               IF #Kamera.text_etiketa = '' THEN
                   #Kamera.text_etiketa := 'NECTENO';   // prazdny text = prazdna pozice!
               END_IF;

               // zapis ZA posledni obsazenou pozici
               #Kamera.idx := 0;
               FOR #i := 5 TO 1 BY -1 DO
                   IF "DB_HMI_recype".fronta[#i].prenaseny_text <> '' THEN
                       #Kamera.idx := #i;
                       EXIT;
                   END_IF;
               END_FOR;

               IF #Kamera.idx < 5 THEN
                   "DB_HMI_recype".fronta[#Kamera.idx + 1].prenaseny_text := #Kamera.text_etiketa;
                   "DB_HMI_recype".fronta[#Kamera.idx + 1].balik_den := #Kamera.balik_den;
                   "DB_HMI_recype".fronta[#Kamera.idx + 1].vyrazeni := #Kamera.vyradit;
               ELSE
                   #Kamera.fronta_plna := TRUE;
               END_IF;
               #Kamera.sber_aktivni := FALSE;
           END_IF;
       END_REGION

       REGION Novy balik pod kamerou - start sberu (az PO zapisu predchoziho)
           IF #Kamera.s2_nabeh THEN
               // citac plat (presunuto ze site 20)
               #zpracovani_dat[1].balik_den := #zpracovani_dat[1].balik_den + 1;
               IF #zpracovani_dat[1].balik_den >= 32000 THEN
                   #zpracovani_dat[1].balik_den := 1;
               END_IF;
               #Kamera.balik_den := #zpracovani_dat[1].balik_den;   // az PO pricteni

               #Kamera.sber_aktivni := TRUE;
               #Kamera.prijato_etiketa := FALSE;
               #Kamera.prijato_folie_l := FALSE;
               #Kamera.prijato_folie_p := FALSE;
               #Kamera.ok_etiketa := FALSE;
               #Kamera.ok_folie_l := FALSE;
               #Kamera.ok_folie_p := FALSE;
               #Kamera.text_etiketa := '';
           END_IF;
       END_REGION
   END_IF;

   REGION Obsazenost fronty pro HMI (pocita se kazdy scan)
       #Kamera.pocet := 0;
       FOR #i := 1 TO 5 DO
           IF "DB_HMI_recype".fronta[#i].prenaseny_text <> '' THEN
               #Kamera.pocet := #Kamera.pocet + 1;
           END_IF;
       END_FOR;
       "DB_HMI_recype".obsazenost_fronty := #Kamera.pocet;
       IF #Kamera.pocet = 0 THEN
           #Kamera.fronta_plna := FALSE;
       END_IF;
   END_REGION
END_REGION

REGION Network 22 (SCL): PŘEPNUTÍ JOBU HORNÍ KAMERY
   // Prepnuti jobu horni kamery podle receptury.
   // Spousti se nabeznou hranou "DB_HMI_recype".ODESLI_dATA (tlacitko Odeslani dat do tiskarny)
   // - soubezne s odeslanim zpravy do tiskarny (OP2).
   // Job 0 v recepture = job neprepinat.

   #Kam_Etiketa_Job.pozadovany := "DB_HMI_recype".recipe.PRG_CAM_etiketa;

   IF "CONTROL_LINE_DB".trig.reset_error_all THEN
       #Kam_Etiketa_Job.chyba := FALSE;
   END_IF;

   CASE #Kam_Etiketa_Job.krok OF
       0:  // ---- klid: cekam na pozadavek ----
           #Kam_Etiketa_Job.aktivni := FALSE;
           "COG_ETIKETA_is3800-ExecuteCommand/JobLoad" := FALSE;
           IF "DB_HMI_recype".ODESLI_dATA AND NOT #Kam_Etiketa_Job.odesli_pamet
               AND #Kam_Etiketa_Job.pozadovany > 0
               AND "COG_ETIKETA_is3800-Online" THEN
               "COG_ETIKETA_is3800-CommandID" := INT_TO_WORD(#Kam_Etiketa_Job.pozadovany);
               #Kam_Etiketa_Job.aktivni := TRUE;
               #Kam_Etiketa_Job.chyba := FALSE;
               #Kam_Etiketa_Job.krok := 10;
           END_IF;

       10: // ---- CommandID uz je venku (predchozi cyklus) -> spustit prikaz ----
           "COG_ETIKETA_is3800-ExecuteCommand/JobLoad" := TRUE;
           #Kam_Etiketa_Job.krok := 20;

       20: // ---- cekam na vysledek ----
           IF "COG_ETIKETA_is3800-CommandCompleted" THEN
               #Kam_Etiketa_Job.krok := 30;
           ELSIF "COG_ETIKETA_is3800-CommandFailed" THEN
               #Kam_Etiketa_Job.chyba := TRUE;
               #Kam_Etiketa_Job.chyba_kod := "COG_ETIKETA_is3800-CommandResultCode";
               #Kam_Etiketa_Job.krok := 30;
           ELSIF #TIMER.TIMER_3.Q THEN
               #Kam_Etiketa_Job.chyba := TRUE;            // kamera neodpovedela
               #Kam_Etiketa_Job.chyba_kod := 16#FFFF;
               #Kam_Etiketa_Job.krok := 30;
           END_IF;

       30: // ---- ukonceni handshake: shodit Execute, pockat az kamera shodi stav ----
           "COG_ETIKETA_is3800-ExecuteCommand/JobLoad" := FALSE;
           IF NOT "COG_ETIKETA_is3800-CommandCompleted"
               AND NOT "COG_ETIKETA_is3800-CommandFailed" THEN
               #Kam_Etiketa_Job.krok := 0;
           END_IF;

       ELSE
           #Kam_Etiketa_Job.krok := 0;
   END_CASE;

   // casovac timeoutu bezi v krocich 10..30
   #TIMER.TIMER_3.TON(IN := #Kam_Etiketa_Job.krok >= 10,
                      PT := #Kam_Etiketa_Job.timeout);
   IF #TIMER.TIMER_3.Q AND #Kam_Etiketa_Job.krok = 30 THEN
       #Kam_Etiketa_Job.krok := 0;                         // pojistka, kdyby kamera stav neshodila
   END_IF;

   #Kam_Etiketa_Job.odesli_pamet := "DB_HMI_recype".ODESLI_dATA;

   // kontrola: v klidu musi job v kamere odpovidat recepture
   #Kam_Etiketa_Job.nesouhlasi := #Kam_Etiketa_Job.krok = 0
   AND #Kam_Etiketa_Job.pozadovany > 0
   AND "COG_ETIKETA_is3800-Online"
   AND WORD_TO_INT("COG_ETIKETA_is3800-Current Job ID") <> #Kam_Etiketa_Job.pozadovany;
END_REGION

REGION Network 23: EXTERNAL_TRIGER
   RUNG wire#powerrail
      { S7_Templates := "SrcType := Int" } EQ_Contact(in1 := #SQCR, in2 := #STEP_5_HOME)
      Contact( "INICIALIZACE_RUN" )
      I_Contact( #TRIG.inicial_ok_op )
      Contact( "AUTOMAT" )
      S_Coil( #HMI.reset_fronty )
      S_Coil( #TRIG.inicial_ok_op )
   END_RUNG
   RUNG wire#powerrail
      Contact( "FirstScan" )
      S_Coil( #HMI.reset_fronty )
      Move(in := 0, out1 => "DB_HMI_recype".obsazenost_fronty, out2 => #zpracovani_dat[1].balik_den)
   END_RUNG
   // the same network as SCL:
   IF (#SQCR = #STEP_5_HOME) AND "INICIALIZACE_RUN" AND NOT #TRIG.inicial_ok_op AND "AUTOMAT" THEN
       #HMI.reset_fronty := TRUE;
       #TRIG.inicial_ok_op := TRUE;
   END_IF;
   IF "FirstScan" THEN
       #HMI.reset_fronty := TRUE;
       "DB_HMI_recype".obsazenost_fronty := 0;
       #zpracovani_dat[1].balik_den := 0;
   END_IF;
END_REGION

REGION Network 24: ETERNAL_TRIGR_INICIAL
   RUNG wire#powerrail
      Contact( "AUTOMAT" )
      { S7_Templates := "SrcType := Int" } GT_Contact(in1 := #SQCR, in2 := #STEP_0)
      { S7_Templates := "SrcType := Int" } LT_Contact(in1 := #SQCR, in2 := #STEP_1000)
      I_Contact( #Kam_Etiketa_Job.aktivni )
      Coil( "COG_ETIKETA_COG_ETIKETA_is3800-TriggerEnable" )
   END_RUNG
   RUNG wire#powerrail
      Contact( "AUTOMAT" )
      { S7_Templates := "SrcType := Int" } GT_Contact(in1 := #SQCR, in2 := #STEP_0)
      { S7_Templates := "SrcType := Int" } LT_Contact(in1 := #SQCR, in2 := #STEP_1000)
      Coil( "COG_FOLIE_L_COG_FOLIE_L_is3800-TriggerEnable" )
   END_RUNG
   RUNG wire#powerrail
      Contact( "AUTOMAT" )
      { S7_Templates := "SrcType := Int" } GT_Contact(in1 := #SQCR, in2 := #STEP_0)
      { S7_Templates := "SrcType := Int" } LT_Contact(in1 := #SQCR, in2 := #STEP_1000)
      Coil( "COG_FOLIE_P_COG_FOLIE_P_is3800-TriggerEnable" )
   END_RUNG
   // the same network as SCL:
   "COG_ETIKETA_COG_ETIKETA_is3800-TriggerEnable" := "AUTOMAT" AND (#SQCR > #STEP_0) AND (#SQCR < #STEP_1000) AND NOT #Kam_Etiketa_Job.aktivni;
   "COG_FOLIE_L_COG_FOLIE_L_is3800-TriggerEnable" := "AUTOMAT" AND (#SQCR > #STEP_0) AND (#SQCR < #STEP_1000);
   "COG_FOLIE_P_COG_FOLIE_P_is3800-TriggerEnable" := "AUTOMAT" AND (#SQCR > #STEP_0) AND (#SQCR < #STEP_1000);
END_REGION

REGION Network 25: hmi
END_REGION

REGION Network 26 (SCL): VYRAZENI MANUAL
   (* #Test_tp_ka12(IN := "DB_Manual".test_vyr,
                 PT := T#500MS);

   "-KA12" := #Test_tp_ka12.Q;

   // testovací bit se sám shodí → každý Modify TRUE = jeden pulz
   IF "DB_Manual".test_vyr THEN
       "DB_Manual".test_vyr := FALSE;
   END_IF; *)
END_REGION
END_FUNCTION_BLOCK

FUNCTION_BLOCK "OP2"   // FB51, LAD
{ S7_Optimized_Access := 'FALSE' }
VERSION : 0.1
   VAR
      CONTROL_MAN : Struct
         B0 : Bool;
         B1 : Bool;
         B2 : Bool;
         B3 : Bool;
         B4 : Bool;
         B5 : Bool;
         B6 : Bool;
         B7 : Bool;
         B8 : Bool;
         B9 : Bool;
         odfuk_1 : Bool;
         odfuk_2 : Bool;
         B12 : Bool;
         B13 : Bool;
         B14 : Bool;
         B15 : Bool;
         B16 : Bool;
         B17 : Bool;
         B18 : Bool;
         B19 : Bool;
         B20 : Bool;
         B21 : Bool;
         B22 : Bool;
         B23 : Bool;
         B24 : Bool;
         B25 : Bool;
         B26 : Bool;
         B27 : Bool;
         B28 : Bool;
         B29 : Bool;
         B30 : Bool;
         B31 : Bool;
      END_STRUCT;
      CONTROL_AUTOMAT : Struct
         connect : Bool;
         send : Bool;
         reciv : Bool;
         trcv : Bool;
         discon : Bool;
         B5 : Bool;
         B6 : Bool;
         B7 : Bool;
         B8 : Bool;
         B9 : Bool;
         B10 : Bool;
         B11 : Bool;
         B12 : Bool;
         B13 : Bool;
         B14 : Bool;
         B15 : Bool;
         B16 : Bool;
         B17 : Bool;
         B18 : Bool;
         B19 : Bool;
         B20 : Bool;
         B21 : Bool;
         B22 : Bool;
         B23 : Bool;
         B24 : Bool;
         B25 : Bool;
         B26 : Bool;
         B27 : Bool;
         B28 : Bool;
         B29 : Bool;
         B30 : Bool;
         B31 : Bool;
      END_STRUCT;
      SENSORS : Struct
         S0 : Bool;
         S1 : Bool;
         S2 : Bool;
         S3 : Bool;
         S4 : Bool;
         S5 : Bool;
         S6 : Bool;
         S7 : Bool;
         S8 : Bool;   // KARUSEL JE NATOČEN PŘÍPRAVKEM A K BRÁNĚ
         S9 : Bool;
         S10 : Bool;
         S11 : Bool;
         S12 : Bool;
         S13 : Bool;
         S14 : Bool;
         S15 : Bool;
         S16 : Bool;
         S17 : Bool;
         S18 : Bool;
         S19 : Bool;
         S20 : Bool;
         S21 : Bool;
         S22 : Bool;
         S23 : Bool;
         S24 : Bool;
         S25 : Bool;
         S26 : Bool;
         S27 : Bool;
         S28 : Bool;
         S29 : Bool;
         S30 : Bool;
         S31 : Bool;
      END_STRUCT;
      SENSORS_1 : Struct
         S0 : Bool;
         S1 : Bool;
         S2 : Bool;
         S3 : Bool;
         S4 : Bool;
         S5 : Bool;
         S6 : Bool;
         S7 : Bool;
         S8 : Bool;
         S9 : Bool;
         S10 : Bool;
         S11 : Bool;
         S12 : Bool;
         S13 : Bool;
         S14 : Bool;
         S15 : Bool;
         S16 : Bool;
         S17 : Bool;
         S18 : Bool;
         S19 : Bool;
         S20 : Bool;
         S21 : Bool;
         S22 : Bool;
         S23 : Bool;
         S24 : Bool;
         S25 : Bool;
         S26 : Bool;
         S27 : Bool;
         S28 : Bool;
         S29 : Bool;
         S30 : Bool;
         S31 : Bool;
      END_STRUCT;
      S_0 : "SENSOR";
      S_1 : "SENSOR";
      S_2 : "SENSOR";
      S_3 : "SENSOR";
      S_4 : "SENSOR";
      S_5 : "SENSOR";
      S_6 : "SENSOR";
      S_7 : "SENSOR";
      S_8 : "SENSOR";
      S_9 : "SENSOR";
      S_10 : "SENSOR";
      S_11 : "SENSOR";
      S_12 : "SENSOR";
      S_13 : "SENSOR";
      S_14 : "SENSOR";
      S_15 : "SENSOR";
      S_16 : "SENSOR";
      M_1 : "MOTOR_CONTROL_BLOCK";
      M_2 : "MOTOR_CONTROL_BLOCK";
      M_3 : "MOTOR_CONTROL_BLOCK";
      SQCR : Int;
      hmi_sqcr : Int;
      TRIG : Struct
         inicial_ok_op : Bool;
         T2 : Bool;
         T3 : Bool;
         T4 : Bool;
         T5 : Bool;
         T6 : Bool;
         T7 : Bool;
         T8 : Bool;
         T9 : Bool;
         T10 : Bool;
         T11 : Bool;
         T12 : Bool;
         T13 : Bool;
         T14 : Bool;
         T15 : Bool;
         T16 : Bool;
         op_1_ready : Bool;
      END_STRUCT;
      MEMOR : Struct
         n_trig_vypnuti : Bool;
         M1 : Bool;
         M2 : Bool;
         M3 : Bool;
         M4 : Bool;
         p_trig_odavacka : Bool;
         M6 : Bool;
         M7 : Bool;
         M8 : Bool;
         M9 : Bool;
         M10 : Bool;
         M11 : Bool;
         RESET_ERROR : Bool;
         M13 : Bool;
         M14 : Bool;
         M15 : Bool;
         SETOVANI_START : Bool;
         M17 : Bool;
         M18 : Bool;
         M19 : Bool;
         M20 : Bool;
         M21 : Bool;
         M22 : Bool;
         M23 : Bool;
         M24 : Bool;
         M25 : Bool;
         M26 : Bool;
         M27 : Bool;
         M28 : Bool;
         M29 : Bool;
         M30 : Bool;
         N_TRIG_SAFETY : Bool;
         M32 : Bool;
         M33 : Bool;
         start_caklu : Bool;
         M35 : Bool;
         M36 : Bool;
         M37 : Bool;
         M38 : Bool;
         M39 : Bool;
         ALARM_GLOBAL : Bool;
         M41 : Bool;
         M42 : Bool;
         M43 : Bool;
         M44 : Bool;
         M45 : Bool;
         M46 : Bool;
         M47 : Bool;
         M48 : Bool;
         M49 : Bool;
         wrong_p_trig : Bool;
         alarm_p_trig : Bool;
         M52 : Bool;
         M53 : Bool;
         M54 : Bool;
         M55 : Bool;
         M56 : Bool;
         M57 : Bool;
         M58 : Bool;
         M59 : Bool;
         M60 : Bool;
         M61 : Bool;
         M62 : Bool;
         M63 : Bool;
      END_STRUCT;
      "TIMER" : Struct
         TIMER_0 : IEC_TIMER;
         TIMER_1 : IEC_TIMER;
         TIMER_2 : IEC_TIMER;
         TIMER_3 : IEC_TIMER;
         TIMER_4 : IEC_TIMER;
         air : IEC_TIMER;
         TIMER_6 : IEC_TIMER;
         TIMER_7 : IEC_TIMER;
      END_STRUCT;
      HMI : Struct
         povoleni_volby_receptu : Bool;
         "svetlo_on/off" : Bool;
         ALARM_VIDITELNOST : Bool;
         hmi_3 : Bool;
         hmi_4 : Bool;
         hmi_5 : Bool;
         hmi_6 : Bool;
         hmi_7 : Bool;
         hmi_8 : Bool;
         hmi_9 : Bool;
         hmi_10 : Bool;
         hmi_11 : Bool;
         hmi_12 : Bool;
         hmi_13 : Bool;
         hmi_14 : Bool;
         hmi_15 : Bool;
      END_STRUCT;
      int_hodnota_zpravy : Word;
      array_do_db AT int_hodnota_zpravy : Array[1..2] of Byte;
      CTRV_LEN : UDInt;
      TCON_Instance : TCON;
      TSEND_Instance : TSEND;
      TRCV_Instance : TRCV;
      TDISCON_Instance : TDISCON;
      Tisk : Struct
         pole2_index_bajt : Int := 14;   // bajt rámce s číslem proměnné
         pole2_index_hodnota : Byte := 16#1;   // číslo proměnné pole 2 (pole 1 = 0)
         datum_chyba : Bool;   // datum přepsáno na XX.XX.XXXX
         pole2_kratky : Bool := true;
         jeden_ramec : Bool;
      END_STRUCT;
   END_VAR
   VAR_TEMP
      DATA : Array[0..255] of Char;
      ARRAY_NULL : Array[1..8] of Bool;
      ARRAY_PRAZDNE : Array[0..255] of Byte;
      j : Int;
      L1 : Int;
      p : Int;
   END_VAR
   VAR CONSTANT
      STEP_0 : Int := 0;
      step_2 : Int := 2;
      STEP_4 : Int := 4;
      STEP_5_HOME : Int := 5;
      STEP_7 : Int := 7;
      STEP_10 : Int := 10;
      STEP_15 : Int := 15;
      STEP_20 : Int := 20;
      STEP_23 : Int := 23;
      STEP_25 : Int := 25;
      STEP_27 : Int := 27;
      STEP_30 : Int := 30;
      STEP_35 : Int := 35;
      STEP_37 : Int := 37;
      STEP_40 : Int := 40;
      STEP_43 : Int := 43;
      STEP_45 : Int := 45;
      STEP_50 : Int := 50;
      STEP_55 : Int := 55;
      STEP_60 : Int := 60;
      STEP_65 : Int := 65;
      STEP_70 : Int := 70;
      STEP_73 : Int := 73;
      STEP_75 : Int := 75;
      STEP_80 : Int := 80;
      STEP_83 : Int := 83;
      STEP_85 : Int := 85;
      STEP_90 : Int := 90;
      STEP_93 : Int := 93;
      STEP_95 : Int := 95;
      STEP_100 : Int := 100;
      STEP_105 : Int := 105;
      STEP_110 : Int := 110;
      STEP_113 : Int := 113;
      STEP_115 : Int := 115;
      STEP_120 : Int := 120;
      STEP_125 : Int := 125;
      STEP_130 : Int := 130;
      STEP_135 : Int := 135;
      STEP_140 : Int := 140;
      STEP_145 : Int := 145;
      STEP_150 : Int := 150;
      STEP_155 : Int := 155;
      STEP_1000 : Int := 1000;
      STEP_1001 : Int := 1001;
      STEP_1002 : Int := 1002;
      STEP_1003 : Int := 1003;
      STEP_1004 : Int := 1004;
      STEP_1005 : Int := 1005;
      STEP_1010 : Int := 1010;
      STEP_1015 : Int := 1015;
      STEP_1020 : Int := 1020;
      STEP_1025 : Int := 1025;
      STEP_3000 : Int := 3000;
      STEP_3005 : Int := 3005;
      STEP_3010 : Int := 3010;
      STEP_3015 : Int := 3015;
      STEP_3020 : Int := 3020;
      STEP_2000 : Int := 2000;
      string_null : String;
      char_null : Char;
      text_kartacek : String := 'Kartacek';
      string_kar_A : String := 'A';
      string_kar_B : String := 'B';
   END_VAR
   VAR_TEMP   // added for the SCL form of the ladder/FBD networks
      _w1 : Bool;
      _w2 : Bool;
      _w3 : Bool;
   END_VAR
BEGIN

REGION Network 1: manuali ovladani reset
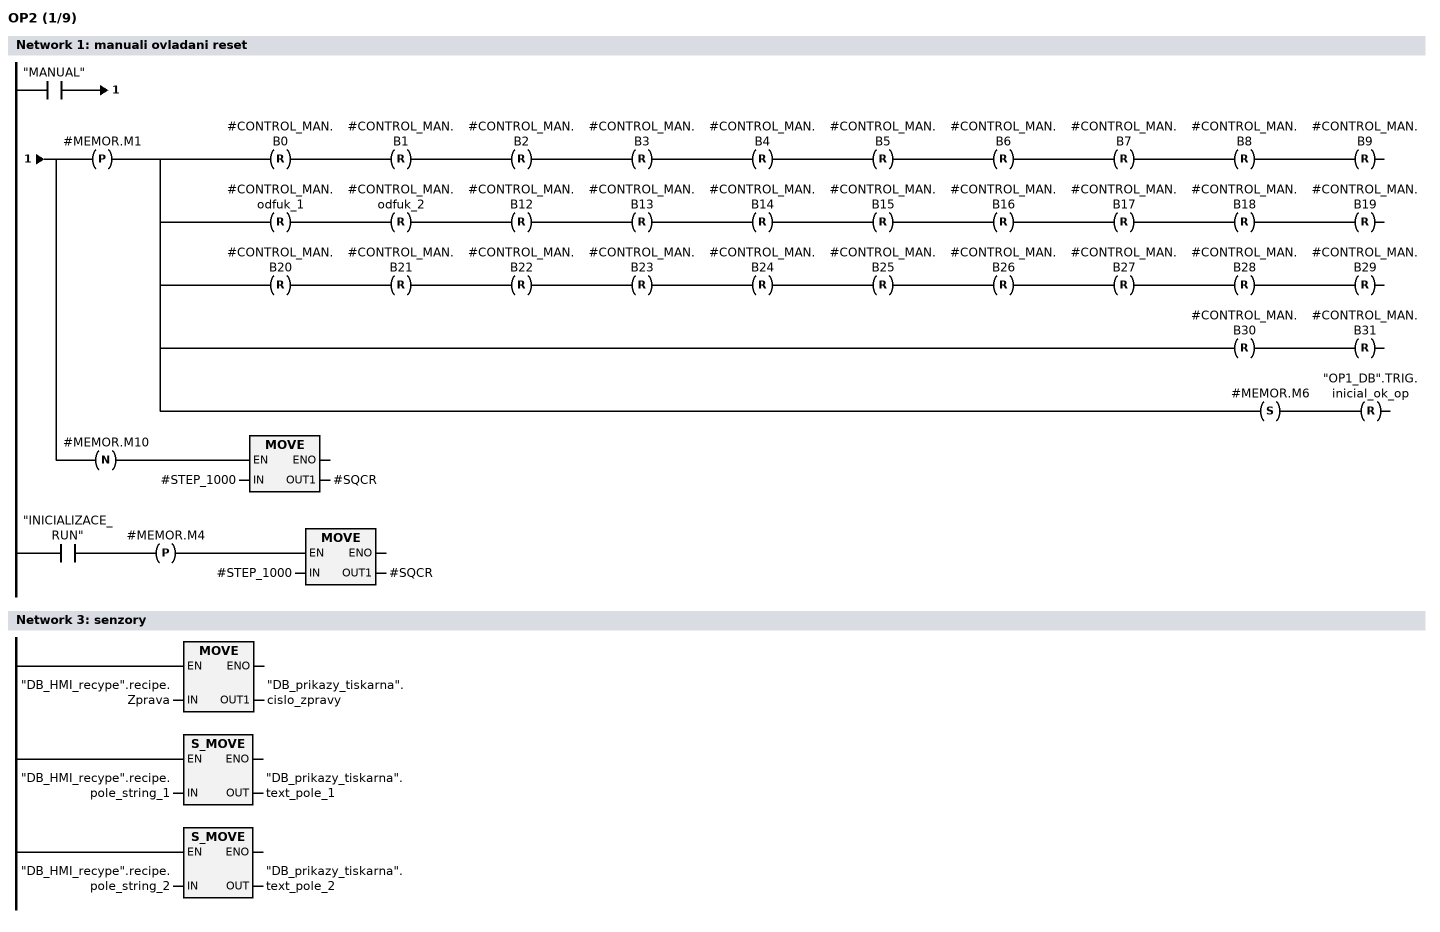
   RUNG wire#powerrail
      Contact( "MANUAL" )
      wire#w1
      P_Trig( #MEMOR.M1 )
      wire#w2
      R_Coil( #CONTROL_MAN.B0 )
      R_Coil( #CONTROL_MAN.B1 )
      R_Coil( #CONTROL_MAN.B2 )
      R_Coil( #CONTROL_MAN.B3 )
      R_Coil( #CONTROL_MAN.B4 )
      R_Coil( #CONTROL_MAN.B5 )
      R_Coil( #CONTROL_MAN.B6 )
      R_Coil( #CONTROL_MAN.B7 )
      R_Coil( #CONTROL_MAN.B8 )
      R_Coil( #CONTROL_MAN.B9 )
   END_RUNG
   RUNG wire#w2
      R_Coil( #CONTROL_MAN.odfuk_1 )
      R_Coil( #CONTROL_MAN.odfuk_2 )
      R_Coil( #CONTROL_MAN.B12 )
      R_Coil( #CONTROL_MAN.B13 )
      R_Coil( #CONTROL_MAN.B14 )
      R_Coil( #CONTROL_MAN.B15 )
      R_Coil( #CONTROL_MAN.B16 )
      R_Coil( #CONTROL_MAN.B17 )
      R_Coil( #CONTROL_MAN.B18 )
      R_Coil( #CONTROL_MAN.B19 )
   END_RUNG
   RUNG wire#w2
      R_Coil( #CONTROL_MAN.B20 )
      R_Coil( #CONTROL_MAN.B21 )
      R_Coil( #CONTROL_MAN.B22 )
      R_Coil( #CONTROL_MAN.B23 )
      R_Coil( #CONTROL_MAN.B24 )
      R_Coil( #CONTROL_MAN.B25 )
      R_Coil( #CONTROL_MAN.B26 )
      R_Coil( #CONTROL_MAN.B27 )
      R_Coil( #CONTROL_MAN.B28 )
      R_Coil( #CONTROL_MAN.B29 )
   END_RUNG
   RUNG wire#w2
      R_Coil( #CONTROL_MAN.B30 )
      R_Coil( #CONTROL_MAN.B31 )
   END_RUNG
   RUNG wire#w2
      S_Coil( #MEMOR.M6 )
      R_Coil( "OP1_DB".TRIG.inicial_ok_op )
   END_RUNG
   RUNG wire#w1
      N_Trig( #MEMOR.M10 )
      Move(in := #STEP_1000, out1 => #SQCR)
   END_RUNG
   RUNG wire#powerrail
      Contact( "INICIALIZACE_RUN" )
      P_Trig( #MEMOR.M4 )
      Move(in := #STEP_1000, out1 => #SQCR)
   END_RUNG
   // the same network as SCL:
   #_w1 := "MANUAL" AND NOT #MEMOR.M1;   // rising edge
   #MEMOR.M1 := "MANUAL";
   IF #_w1 THEN
       #CONTROL_MAN.B0 := FALSE;
       #CONTROL_MAN.B1 := FALSE;
       #CONTROL_MAN.B2 := FALSE;
       #CONTROL_MAN.B3 := FALSE;
       #CONTROL_MAN.B4 := FALSE;
       #CONTROL_MAN.B5 := FALSE;
       #CONTROL_MAN.B6 := FALSE;
       #CONTROL_MAN.B7 := FALSE;
       #CONTROL_MAN.B8 := FALSE;
       #CONTROL_MAN.B9 := FALSE;
       #CONTROL_MAN.odfuk_1 := FALSE;
       #CONTROL_MAN.odfuk_2 := FALSE;
       #CONTROL_MAN.B12 := FALSE;
       #CONTROL_MAN.B13 := FALSE;
       #CONTROL_MAN.B14 := FALSE;
       #CONTROL_MAN.B15 := FALSE;
       #CONTROL_MAN.B16 := FALSE;
       #CONTROL_MAN.B17 := FALSE;
       #CONTROL_MAN.B18 := FALSE;
       #CONTROL_MAN.B19 := FALSE;
       #CONTROL_MAN.B20 := FALSE;
       #CONTROL_MAN.B21 := FALSE;
       #CONTROL_MAN.B22 := FALSE;
       #CONTROL_MAN.B23 := FALSE;
       #CONTROL_MAN.B24 := FALSE;
       #CONTROL_MAN.B25 := FALSE;
       #CONTROL_MAN.B26 := FALSE;
       #CONTROL_MAN.B27 := FALSE;
       #CONTROL_MAN.B28 := FALSE;
       #CONTROL_MAN.B29 := FALSE;
       #CONTROL_MAN.B30 := FALSE;
       #CONTROL_MAN.B31 := FALSE;
       #MEMOR.M6 := TRUE;
       "OP1_DB".TRIG.inicial_ok_op := FALSE;
   END_IF;
   #_w2 := NOT "MANUAL" AND #MEMOR.M10;   // falling edge
   #MEMOR.M10 := "MANUAL";
   IF #_w2 THEN #SQCR := #STEP_1000; END_IF;
   #_w3 := "INICIALIZACE_RUN" AND NOT #MEMOR.M4;   // rising edge
   #MEMOR.M4 := "INICIALIZACE_RUN";
   IF #_w3 THEN #SQCR := #STEP_1000; END_IF;
END_REGION

REGION Network 2: alarmy
END_REGION

REGION Network 3: senzory
   RUNG wire#powerrail
      Move(in := "DB_HMI_recype".recipe.Zprava, out1 => "DB_prikazy_tiskarna".cislo_zpravy)
   END_RUNG
   RUNG wire#powerrail
      S_Move(in := "DB_HMI_recype".recipe.pole_string_1, out => "DB_prikazy_tiskarna".text_pole_1)
   END_RUNG
   RUNG wire#powerrail
      S_Move(in := "DB_HMI_recype".recipe.pole_string_2, out => "DB_prikazy_tiskarna".text_pole_2)
   END_RUNG
   // the same network as SCL:
   "DB_prikazy_tiskarna".cislo_zpravy := "DB_HMI_recype".recipe.Zprava;
   "DB_prikazy_tiskarna".text_pole_1 := "DB_HMI_recype".recipe.pole_string_1;
   "DB_prikazy_tiskarna".text_pole_2 := "DB_HMI_recype".recipe.pole_string_2;
END_REGION

REGION Network 4 (SCL): tiskarna_zpracovani_dat


   #int_hodnota_zpravy := "DB_prikazy_tiskarna".cislo_zpravy;


   //"DB_prikazy_tiskarna".byte_2 := INT_TO_CHAR( "DB_prikazy_tiskarna".cislo_zpravy);
   "DB_prikazy_tiskarna".byte_1 := #array_do_db[1] + 48;
   "DB_prikazy_tiskarna".byte_2 := #array_do_db[2] + 48;


   "DB_prikazy_tiskarna".task[3, 26] := "DB_prikazy_tiskarna".byte_1;
   "DB_prikazy_tiskarna".task[3, 27] := "DB_prikazy_tiskarna".byte_2;











   "DB_prikazy_tiskarna".task[4, 17] := "DB_prikazy_tiskarna".text_pole_1[1];
   "DB_prikazy_tiskarna".task[4, 18] := "DB_prikazy_tiskarna".text_pole_1[2];
   "DB_prikazy_tiskarna".task[4, 19] := "DB_prikazy_tiskarna".text_pole_1[3];
   "DB_prikazy_tiskarna".task[4, 20] := "DB_prikazy_tiskarna".text_pole_1[4];
   "DB_prikazy_tiskarna".task[4, 21] := "DB_prikazy_tiskarna".text_pole_1[5];
   "DB_prikazy_tiskarna".task[4, 22] := "DB_prikazy_tiskarna".text_pole_1[6];
   "DB_prikazy_tiskarna".task[4, 23] := "DB_prikazy_tiskarna".text_pole_1[7];
   "DB_prikazy_tiskarna".task[4, 24] := "DB_prikazy_tiskarna".text_pole_1[8];
   "DB_prikazy_tiskarna".task[4, 25] := "DB_prikazy_tiskarna".text_pole_1[9];
   "DB_prikazy_tiskarna".task[4, 26] := "DB_prikazy_tiskarna".text_pole_1[10];
   "DB_prikazy_tiskarna".task[4, 27] := "DB_prikazy_tiskarna".text_pole_1[11];
   "DB_prikazy_tiskarna".task[4, 28] := "DB_prikazy_tiskarna".text_pole_1[12];
   "DB_prikazy_tiskarna".task[4, 29] := "DB_prikazy_tiskarna".text_pole_1[13];
   "DB_prikazy_tiskarna".task[4, 30] := "DB_prikazy_tiskarna".text_pole_1[14];
   "DB_prikazy_tiskarna".task[4, 31] := "DB_prikazy_tiskarna".text_pole_1[15];
   "DB_prikazy_tiskarna".task[4, 32] := "DB_prikazy_tiskarna".text_pole_1[16];
   "DB_prikazy_tiskarna".task[4, 33] := "DB_prikazy_tiskarna".text_pole_1[17];
   "DB_prikazy_tiskarna".task[4, 34] := "DB_prikazy_tiskarna".text_pole_1[18];
   "DB_prikazy_tiskarna".task[4, 35] := "DB_prikazy_tiskarna".text_pole_1[19];
   "DB_prikazy_tiskarna".task[4, 36] := "DB_prikazy_tiskarna".text_pole_1[20];
   "DB_prikazy_tiskarna".task[4, 37] := "DB_prikazy_tiskarna".text_pole_1[21];
   "DB_prikazy_tiskarna".task[4, 38] := "DB_prikazy_tiskarna".text_pole_1[22];
   "DB_prikazy_tiskarna".task[4, 39] := "DB_prikazy_tiskarna".text_pole_1[23];
   "DB_prikazy_tiskarna".task[4, 40] := "DB_prikazy_tiskarna".text_pole_1[24];
   "DB_prikazy_tiskarna".task[4, 41] := "DB_prikazy_tiskarna".text_pole_1[25];
   "DB_prikazy_tiskarna".task[4, 42] := "DB_prikazy_tiskarna".text_pole_1[26];
   "DB_prikazy_tiskarna".task[4, 43] := "DB_prikazy_tiskarna".text_pole_1[27];
   "DB_prikazy_tiskarna".task[4, 44] := "DB_prikazy_tiskarna".text_pole_1[28];
   "DB_prikazy_tiskarna".task[4, 45] := "DB_prikazy_tiskarna".text_pole_1[29];
   "DB_prikazy_tiskarna".task[4, 46] := "DB_prikazy_tiskarna".text_pole_1[30];






   IF "DB_HMI_recype".recipe.pole_string_2[3] <> '.' OR "DB_HMI_recype".recipe.pole_string_2[6] <> '.' THEN
       "DB_HMI_recype".recipe.pole_string_2 := 'XX.XX.XXXX';
   END_IF;



   // ===================== POLE 2 - DATUM SPOTREBY (radek 5) =====================
   // Samostatny ramec CF stejny jako pole 1 (radek 4), lisi se cislem promenne,
   // delkou textu a obsahem. Odesila se v kroku 130 (ADRESACE_POLE = 5).

   // chybne datum (prepsane na XX) -> priznak pro alarm / vyrazeni
   #Tisk.datum_chyba := "DB_HMI_recype".recipe.pole_string_2 = 'XX.XX.XXXX';

   // hlavicka ramce = kopie hlavicky pole 1 (bajty 0..16)
   FOR #j := 0 TO 16 DO
       "DB_prikazy_tiskarna".task[5, #j] := "DB_prikazy_tiskarna".task[4, #j];
   END_FOR;

   // cislo promenne pole 2 - bajt nastavitelny (12/13/14), overit na tiskarne
   IF #Tisk.pole2_index_bajt >= 12 AND #Tisk.pole2_index_bajt <= 14 THEN
       "DB_prikazy_tiskarna".task[5, #Tisk.pole2_index_bajt] := #Tisk.pole2_index_hodnota;
   END_IF;

   // datum - vzdy 10 znaku (DD.MM.RRRR nebo XX.XX.XXXX)
   "DB_prikazy_tiskarna".task[5, 17] := "DB_prikazy_tiskarna".text_pole_2[1];
   "DB_prikazy_tiskarna".task[5, 18] := "DB_prikazy_tiskarna".text_pole_2[2];
   "DB_prikazy_tiskarna".task[5, 19] := "DB_prikazy_tiskarna".text_pole_2[3];
   "DB_prikazy_tiskarna".task[5, 20] := "DB_prikazy_tiskarna".text_pole_2[4];
   "DB_prikazy_tiskarna".task[5, 21] := "DB_prikazy_tiskarna".text_pole_2[5];
   "DB_prikazy_tiskarna".task[5, 22] := "DB_prikazy_tiskarna".text_pole_2[6];
   "DB_prikazy_tiskarna".task[5, 23] := "DB_prikazy_tiskarna".text_pole_2[7];
   "DB_prikazy_tiskarna".task[5, 24] := "DB_prikazy_tiskarna".text_pole_2[8];
   "DB_prikazy_tiskarna".task[5, 25] := "DB_prikazy_tiskarna".text_pole_2[9];
   "DB_prikazy_tiskarna".task[5, 26] := "DB_prikazy_tiskarna".text_pole_2[10];

   IF #Tisk.pole2_kratky THEN
       // --- 10 znaku: upravit delky v hlavicce ---
       "DB_prikazy_tiskarna".task[5, 5] := 16#28;   // delka ramce od bajtu 6 = 40
       "DB_prikazy_tiskarna".task[5, 8] := 16#00;
       "DB_prikazy_tiskarna".task[5, 9] := 16#24;   // delka dat prikazu od bajtu 10 = 36
       "DB_prikazy_tiskarna".task[5, 15] := 16#00;
       "DB_prikazy_tiskarna".task[5, 16] := 16#0A;   // delka textu = 10 znaku
       // za datem 19 x 00 (bajty 27..45), dal nic
       FOR #j := 27 TO 65 DO
           "DB_prikazy_tiskarna".task[5, #j] := 16#00;
       END_FOR;
   ELSE
       // --- 30 znaku (puvodni varianta): delky z hlavicky pole 1, doplnit mezerami ---
       FOR #j := 27 TO 46 DO
           "DB_prikazy_tiskarna".task[5, #j] := 16#20;
       END_FOR;
       FOR #j := 47 TO 65 DO
           "DB_prikazy_tiskarna".task[5, #j] := 16#00;
       END_FOR;
   END_IF;

   // ===== OBE POLE V JEDNOM RAMCI CF: 20 promennych, delka 1 bajt =====
   IF #Tisk.jeden_ramec THEN
       #L1 := LEN("DB_prikazy_tiskarna".text_pole_1);
       IF #L1 > 30 THEN
           #L1 := 30;
       END_IF;

       FOR #j := 15 TO 120 DO
           "DB_prikazy_tiskarna".task[4, #j] := 16#00;
       END_FOR;

       // promenna 1: delka (1 bajt) + Puvod
       "DB_prikazy_tiskarna".task[4, 16] := INT_TO_BYTE(#L1);
       FOR #j := 1 TO #L1 DO
           "DB_prikazy_tiskarna".task[4, 16 + #j] := "DB_prikazy_tiskarna".text_pole_1[#j];
       END_FOR;
       #p := 17 + #L1;

       // promenna 2: delka (1 bajt) + datum
       "DB_prikazy_tiskarna".task[4, #p] := 16#0A;
       FOR #j := 1 TO 10 DO
           "DB_prikazy_tiskarna".task[4, #p + #j] := "DB_prikazy_tiskarna".text_pole_2[#j];
       END_FOR;
       #p := #p + 11;

       // promenne 3..20 prazdne = 18 x 00 (uz vycisteno)
       #p := #p + 18;

       "DB_prikazy_tiskarna".task[4, 4] := 16#00;
       "DB_prikazy_tiskarna".task[4, 5] := INT_TO_BYTE(#p - 6);
       "DB_prikazy_tiskarna".task[4, 8] := 16#00;
       "DB_prikazy_tiskarna".task[4, 9] := INT_TO_BYTE(#p - 10);
   END_IF;
END_REGION

REGION Network 5: příkazy k odeslání z bafru
   // 2 = STOP TISKU
   // 3 = VÝBĚR ZPRÁVY
   // 6 = NASTAVENÍ NEBAFROVÁNÍ A SMAZÁNÍ PŘEDEŠLÍCH DAT
   // 4 = ZAPSÁNÍ DO VARIABILNÍHO POLE 1
   // 5 = ZAPSÁNÍ DO VARIABILNÍHO POLE 2
   // 1 = START TISKU
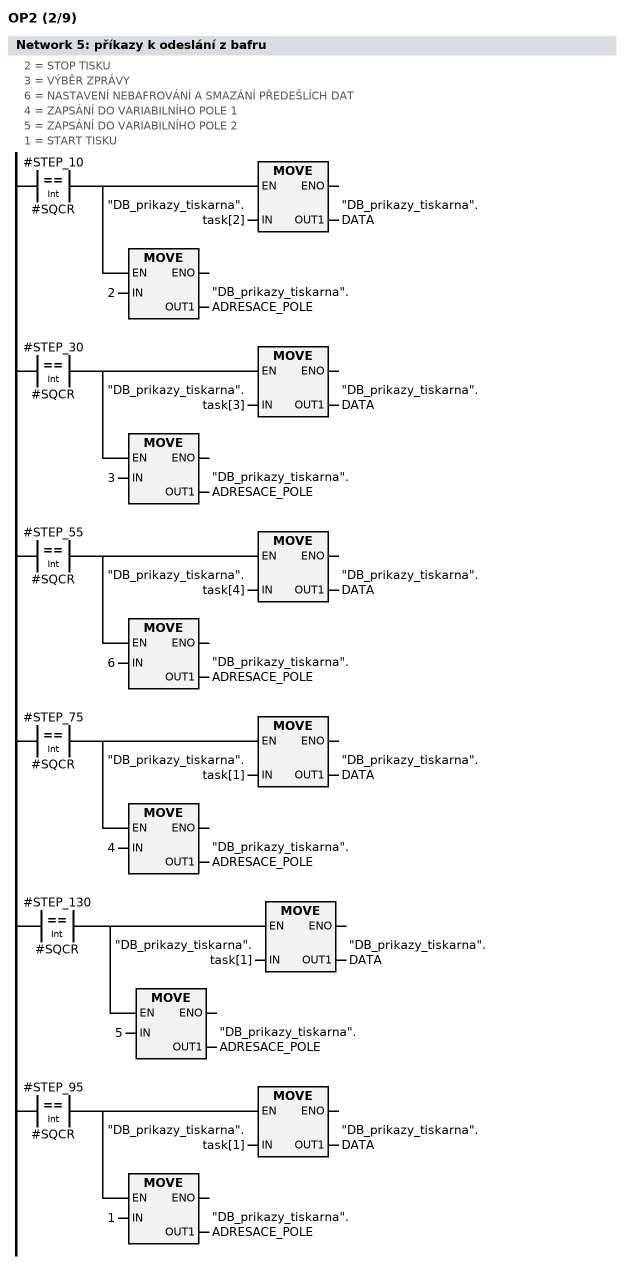
   RUNG wire#powerrail
      { S7_Templates := "SrcType := Int" } EQ_Contact(in1 := #STEP_10, in2 := #SQCR)
      wire#w1
      Move(in := "DB_prikazy_tiskarna".task[2], out1 => "DB_prikazy_tiskarna".DATA)
   END_RUNG
   RUNG wire#w1
      Move(in := 2, out1 => "DB_prikazy_tiskarna".ADRESACE_POLE)
   END_RUNG
   RUNG wire#powerrail
      { S7_Templates := "SrcType := Int" } EQ_Contact(in1 := #STEP_30, in2 := #SQCR)
      wire#w2
      Move(in := "DB_prikazy_tiskarna".task[3], out1 => "DB_prikazy_tiskarna".DATA)
   END_RUNG
   RUNG wire#w2
      Move(in := 3, out1 => "DB_prikazy_tiskarna".ADRESACE_POLE)
   END_RUNG
   RUNG wire#powerrail
      { S7_Templates := "SrcType := Int" } EQ_Contact(in1 := #STEP_55, in2 := #SQCR)
      wire#w3
      Move(in := "DB_prikazy_tiskarna".task[4], out1 => "DB_prikazy_tiskarna".DATA)
   END_RUNG
   RUNG wire#w3
      Move(in := 6, out1 => "DB_prikazy_tiskarna".ADRESACE_POLE)
   END_RUNG
   RUNG wire#powerrail
      { S7_Templates := "SrcType := Int" } EQ_Contact(in1 := #STEP_75, in2 := #SQCR)
      wire#w4
      Move(in := "DB_prikazy_tiskarna".task[1], out1 => "DB_prikazy_tiskarna".DATA)
   END_RUNG
   RUNG wire#w4
      Move(in := 4, out1 => "DB_prikazy_tiskarna".ADRESACE_POLE)
   END_RUNG
   RUNG wire#powerrail
      { S7_Templates := "SrcType := Int" } EQ_Contact(in1 := #STEP_130, in2 := #SQCR)
      wire#w5
      Move(in := "DB_prikazy_tiskarna".task[1], out1 => "DB_prikazy_tiskarna".DATA)
   END_RUNG
   RUNG wire#w5
      Move(in := 5, out1 => "DB_prikazy_tiskarna".ADRESACE_POLE)
   END_RUNG
   RUNG wire#powerrail
      { S7_Templates := "SrcType := Int" } EQ_Contact(in1 := #STEP_95, in2 := #SQCR)
      wire#w6
      Move(in := "DB_prikazy_tiskarna".task[1], out1 => "DB_prikazy_tiskarna".DATA)
   END_RUNG
   RUNG wire#w6
      Move(in := 1, out1 => "DB_prikazy_tiskarna".ADRESACE_POLE)
   END_RUNG
   // the same network as SCL:
   IF #STEP_10 = #SQCR THEN
       "DB_prikazy_tiskarna".DATA := "DB_prikazy_tiskarna".task[2];
       "DB_prikazy_tiskarna".ADRESACE_POLE := 2;
   END_IF;
   IF #STEP_30 = #SQCR THEN
       "DB_prikazy_tiskarna".DATA := "DB_prikazy_tiskarna".task[3];
       "DB_prikazy_tiskarna".ADRESACE_POLE := 3;
   END_IF;
   IF #STEP_55 = #SQCR THEN
       "DB_prikazy_tiskarna".DATA := "DB_prikazy_tiskarna".task[4];
       "DB_prikazy_tiskarna".ADRESACE_POLE := 6;
   END_IF;
   IF #STEP_75 = #SQCR THEN
       "DB_prikazy_tiskarna".DATA := "DB_prikazy_tiskarna".task[1];
       "DB_prikazy_tiskarna".ADRESACE_POLE := 4;
   END_IF;
   IF #STEP_130 = #SQCR THEN
       "DB_prikazy_tiskarna".DATA := "DB_prikazy_tiskarna".task[1];
       "DB_prikazy_tiskarna".ADRESACE_POLE := 5;
   END_IF;
   IF #STEP_95 = #SQCR THEN
       "DB_prikazy_tiskarna".DATA := "DB_prikazy_tiskarna".task[1];
       "DB_prikazy_tiskarna".ADRESACE_POLE := 1;
   END_IF;
END_REGION

REGION Network 6: CONTROL BLOCK tiskarna
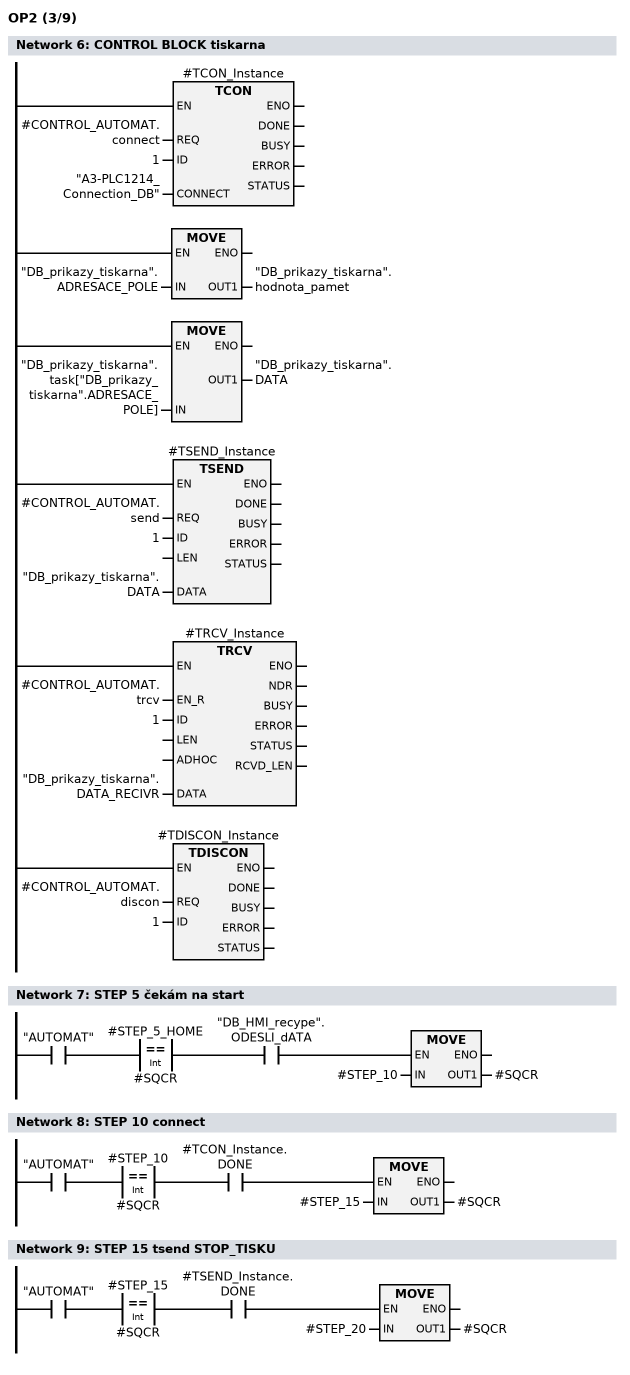
   #TCON_Instance(REQ := #CONTROL_AUTOMAT.connect, ID := 1, CONNECT := "A3-PLC1214_Connection_DB");   // TCON
   "DB_prikazy_tiskarna".hodnota_pamet := "DB_prikazy_tiskarna".ADRESACE_POLE;
   "DB_prikazy_tiskarna".DATA := "DB_prikazy_tiskarna".task["DB_prikazy_tiskarna".ADRESACE_POLE];
   #TSEND_Instance(REQ := #CONTROL_AUTOMAT.send, ID := 1, DATA := "DB_prikazy_tiskarna".DATA);   // TSEND
   #TRCV_Instance(EN_R := #CONTROL_AUTOMAT.trcv, ID := 1, DATA := "DB_prikazy_tiskarna".DATA_RECIVR);   // TRCV
   #TDISCON_Instance(REQ := #CONTROL_AUTOMAT.discon, ID := 1);   // TDISCON
END_REGION

REGION Network 7: STEP 5 čekám na start
   RUNG wire#powerrail
      Contact( "AUTOMAT" )
      { S7_Templates := "SrcType := Int" } EQ_Contact(in1 := #STEP_5_HOME, in2 := #SQCR)
      Contact( "DB_HMI_recype".ODESLI_dATA )
      Move(in := #STEP_10, out1 => #SQCR)
   END_RUNG
   // the same network as SCL:
   IF "AUTOMAT" AND (#STEP_5_HOME = #SQCR) AND "DB_HMI_recype".ODESLI_dATA THEN #SQCR := #STEP_10; END_IF;
END_REGION

REGION Network 8: STEP 10 connect
   RUNG wire#powerrail
      Contact( "AUTOMAT" )
      { S7_Templates := "SrcType := Int" } EQ_Contact(in1 := #STEP_10, in2 := #SQCR)
      Contact( #TCON_Instance.DONE )
      Move(in := #STEP_15, out1 => #SQCR)
   END_RUNG
   // the same network as SCL:
   IF "AUTOMAT" AND (#STEP_10 = #SQCR) AND #TCON_Instance.DONE THEN #SQCR := #STEP_15; END_IF;
END_REGION

REGION Network 9: STEP 15 tsend STOP_TISKU
   RUNG wire#powerrail
      Contact( "AUTOMAT" )
      { S7_Templates := "SrcType := Int" } EQ_Contact(in1 := #STEP_15, in2 := #SQCR)
      Contact( #TSEND_Instance.DONE )
      Move(in := #STEP_20, out1 => #SQCR)
   END_RUNG
   // the same network as SCL:
   IF "AUTOMAT" AND (#STEP_15 = #SQCR) AND #TSEND_Instance.DONE THEN #SQCR := #STEP_20; END_IF;
END_REGION

REGION Network 10: STEP 20 odpověď
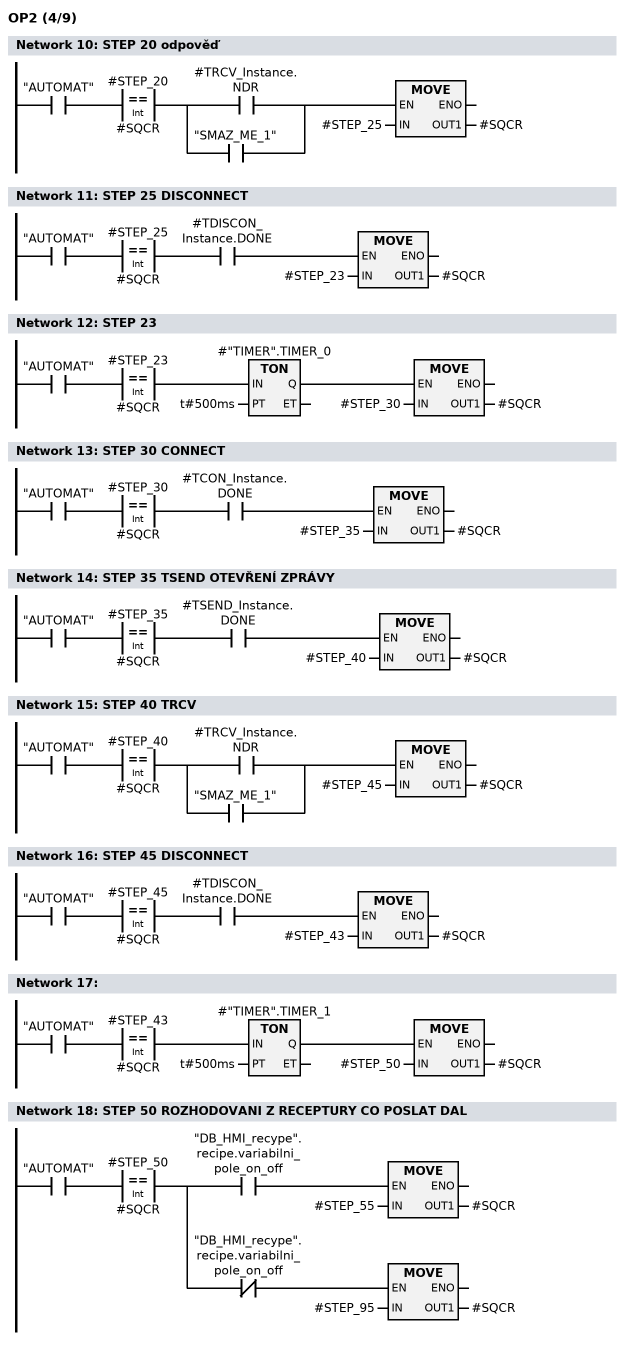
   RUNG wire#powerrail
      Contact( "AUTOMAT" )
      { S7_Templates := "SrcType := Int" } EQ_Contact(in1 := #STEP_20, in2 := #SQCR)
      wire#w1
      Contact( #TRCV_Instance.NDR )
      wire#w2
      Move(in := #STEP_25, out1 => #SQCR)
   END_RUNG
   RUNG wire#w1
      Contact( "SMAZ_ME_1" )
   END_RUNG wire#w2
   // the same network as SCL:
   IF "AUTOMAT" AND (#STEP_20 = #SQCR) AND (#TRCV_Instance.NDR OR "SMAZ_ME_1") THEN
       #SQCR := #STEP_25;
   END_IF;
END_REGION

REGION Network 11: STEP 25 DISCONNECT
   RUNG wire#powerrail
      Contact( "AUTOMAT" )
      { S7_Templates := "SrcType := Int" } EQ_Contact(in1 := #STEP_25, in2 := #SQCR)
      Contact( #TDISCON_Instance.DONE )
      Move(in := #STEP_23, out1 => #SQCR)
   END_RUNG
   // the same network as SCL:
   IF "AUTOMAT" AND (#STEP_25 = #SQCR) AND #TDISCON_Instance.DONE THEN #SQCR := #STEP_23; END_IF;
END_REGION

REGION Network 12: STEP 23
   #"TIMER".TIMER_0.TON(IN := "AUTOMAT" AND (#STEP_23 = #SQCR), PT := t#500ms);
   IF #"TIMER".TIMER_0.Q THEN #SQCR := #STEP_30; END_IF;
END_REGION

REGION Network 13: STEP 30 CONNECT
   RUNG wire#powerrail
      Contact( "AUTOMAT" )
      { S7_Templates := "SrcType := Int" } EQ_Contact(in1 := #STEP_30, in2 := #SQCR)
      Contact( #TCON_Instance.DONE )
      Move(in := #STEP_35, out1 => #SQCR)
   END_RUNG
   // the same network as SCL:
   IF "AUTOMAT" AND (#STEP_30 = #SQCR) AND #TCON_Instance.DONE THEN #SQCR := #STEP_35; END_IF;
END_REGION

REGION Network 14: STEP 35 TSEND OTEVŘENÍ ZPRÁVY
   RUNG wire#powerrail
      Contact( "AUTOMAT" )
      { S7_Templates := "SrcType := Int" } EQ_Contact(in1 := #STEP_35, in2 := #SQCR)
      Contact( #TSEND_Instance.DONE )
      Move(in := #STEP_40, out1 => #SQCR)
   END_RUNG
   // the same network as SCL:
   IF "AUTOMAT" AND (#STEP_35 = #SQCR) AND #TSEND_Instance.DONE THEN #SQCR := #STEP_40; END_IF;
END_REGION

REGION Network 15: STEP 40 TRCV
   RUNG wire#powerrail
      Contact( "AUTOMAT" )
      { S7_Templates := "SrcType := Int" } EQ_Contact(in1 := #STEP_40, in2 := #SQCR)
      wire#w1
      Contact( #TRCV_Instance.NDR )
      wire#w2
      Move(in := #STEP_45, out1 => #SQCR)
   END_RUNG
   RUNG wire#w1
      Contact( "SMAZ_ME_1" )
   END_RUNG wire#w2
   // the same network as SCL:
   IF "AUTOMAT" AND (#STEP_40 = #SQCR) AND (#TRCV_Instance.NDR OR "SMAZ_ME_1") THEN
       #SQCR := #STEP_45;
   END_IF;
END_REGION

REGION Network 16: STEP 45 DISCONNECT
   RUNG wire#powerrail
      Contact( "AUTOMAT" )
      { S7_Templates := "SrcType := Int" } EQ_Contact(in1 := #STEP_45, in2 := #SQCR)
      Contact( #TDISCON_Instance.DONE )
      Move(in := #STEP_43, out1 => #SQCR)
   END_RUNG
   // the same network as SCL:
   IF "AUTOMAT" AND (#STEP_45 = #SQCR) AND #TDISCON_Instance.DONE THEN #SQCR := #STEP_43; END_IF;
END_REGION

REGION Network 17
   #"TIMER".TIMER_1.TON(IN := "AUTOMAT" AND (#STEP_43 = #SQCR), PT := t#500ms);
   IF #"TIMER".TIMER_1.Q THEN #SQCR := #STEP_50; END_IF;
END_REGION

REGION Network 18: STEP 50 ROZHODOVANI Z RECEPTURY CO POSLAT DAL
   RUNG wire#powerrail
      Contact( "AUTOMAT" )
      { S7_Templates := "SrcType := Int" } EQ_Contact(in1 := #STEP_50, in2 := #SQCR)
      wire#w1
      Contact( "DB_HMI_recype".recipe.variabilni_pole_on_off )
      Move(in := #STEP_55, out1 => #SQCR)
   END_RUNG
   RUNG wire#w1
      I_Contact( "DB_HMI_recype".recipe.variabilni_pole_on_off )
      Move(in := #STEP_95, out1 => #SQCR)
   END_RUNG
   // the same network as SCL:
   #_w1 := "AUTOMAT" AND (#STEP_50 = #SQCR);
   IF #_w1 AND "DB_HMI_recype".recipe.variabilni_pole_on_off THEN #SQCR := #STEP_55; END_IF;
   IF #_w1 AND NOT "DB_HMI_recype".recipe.variabilni_pole_on_off THEN #SQCR := #STEP_95; END_IF;
END_REGION

REGION Network 19: STEP 55 CONNECT
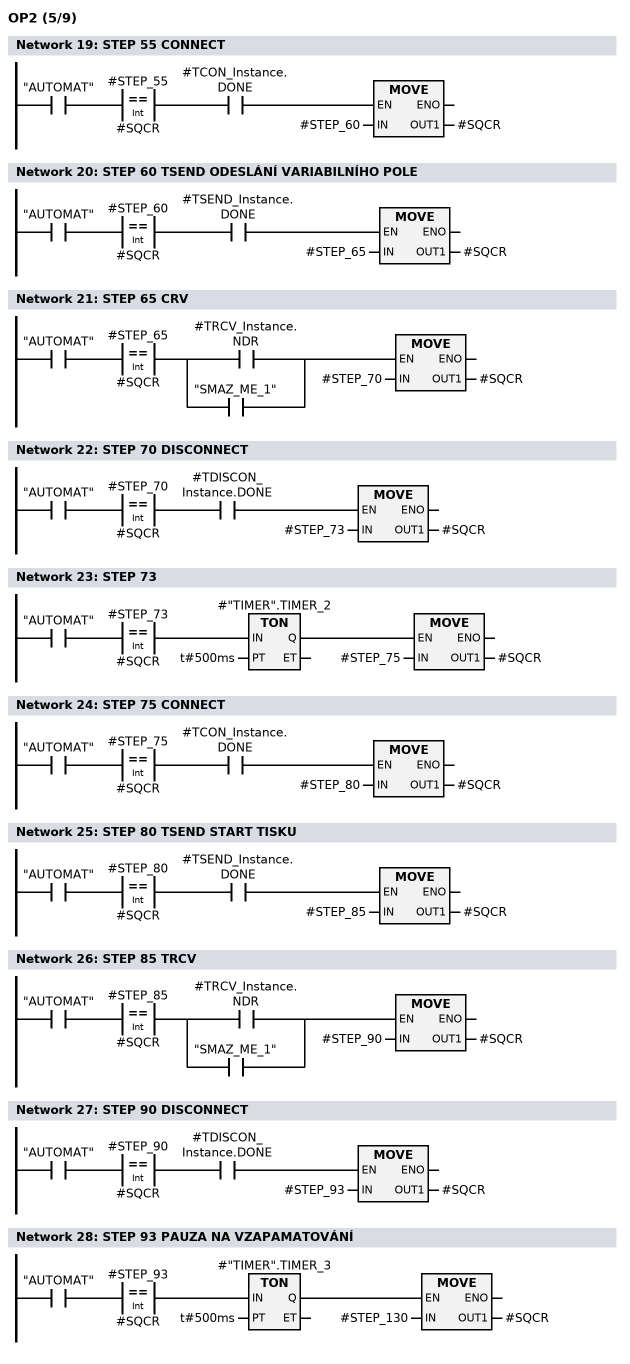
   RUNG wire#powerrail
      Contact( "AUTOMAT" )
      { S7_Templates := "SrcType := Int" } EQ_Contact(in1 := #STEP_55, in2 := #SQCR)
      Contact( #TCON_Instance.DONE )
      Move(in := #STEP_60, out1 => #SQCR)
   END_RUNG
   // the same network as SCL:
   IF "AUTOMAT" AND (#STEP_55 = #SQCR) AND #TCON_Instance.DONE THEN #SQCR := #STEP_60; END_IF;
END_REGION

REGION Network 20: STEP 60 TSEND ODESLÁNÍ VARIABILNÍHO POLE
   RUNG wire#powerrail
      Contact( "AUTOMAT" )
      { S7_Templates := "SrcType := Int" } EQ_Contact(in1 := #STEP_60, in2 := #SQCR)
      Contact( #TSEND_Instance.DONE )
      Move(in := #STEP_65, out1 => #SQCR)
   END_RUNG
   // the same network as SCL:
   IF "AUTOMAT" AND (#STEP_60 = #SQCR) AND #TSEND_Instance.DONE THEN #SQCR := #STEP_65; END_IF;
END_REGION

REGION Network 21: STEP 65 CRV
   RUNG wire#powerrail
      Contact( "AUTOMAT" )
      { S7_Templates := "SrcType := Int" } EQ_Contact(in1 := #STEP_65, in2 := #SQCR)
      wire#w1
      Contact( #TRCV_Instance.NDR )
      wire#w2
      Move(in := #STEP_70, out1 => #SQCR)
   END_RUNG
   RUNG wire#w1
      Contact( "SMAZ_ME_1" )
   END_RUNG wire#w2
   // the same network as SCL:
   IF "AUTOMAT" AND (#STEP_65 = #SQCR) AND (#TRCV_Instance.NDR OR "SMAZ_ME_1") THEN
       #SQCR := #STEP_70;
   END_IF;
END_REGION

REGION Network 22: STEP 70 DISCONNECT
   RUNG wire#powerrail
      Contact( "AUTOMAT" )
      { S7_Templates := "SrcType := Int" } EQ_Contact(in1 := #STEP_70, in2 := #SQCR)
      Contact( #TDISCON_Instance.DONE )
      Move(in := #STEP_73, out1 => #SQCR)
   END_RUNG
   // the same network as SCL:
   IF "AUTOMAT" AND (#STEP_70 = #SQCR) AND #TDISCON_Instance.DONE THEN #SQCR := #STEP_73; END_IF;
END_REGION

REGION Network 23: STEP 73
   #"TIMER".TIMER_2.TON(IN := "AUTOMAT" AND (#STEP_73 = #SQCR), PT := t#500ms);
   IF #"TIMER".TIMER_2.Q THEN #SQCR := #STEP_75; END_IF;
END_REGION

REGION Network 24: STEP 75 CONNECT
   RUNG wire#powerrail
      Contact( "AUTOMAT" )
      { S7_Templates := "SrcType := Int" } EQ_Contact(in1 := #STEP_75, in2 := #SQCR)
      Contact( #TCON_Instance.DONE )
      Move(in := #STEP_80, out1 => #SQCR)
   END_RUNG
   // the same network as SCL:
   IF "AUTOMAT" AND (#STEP_75 = #SQCR) AND #TCON_Instance.DONE THEN #SQCR := #STEP_80; END_IF;
END_REGION

REGION Network 25: STEP 80 TSEND START TISKU
   RUNG wire#powerrail
      Contact( "AUTOMAT" )
      { S7_Templates := "SrcType := Int" } EQ_Contact(in1 := #STEP_80, in2 := #SQCR)
      Contact( #TSEND_Instance.DONE )
      Move(in := #STEP_85, out1 => #SQCR)
   END_RUNG
   // the same network as SCL:
   IF "AUTOMAT" AND (#STEP_80 = #SQCR) AND #TSEND_Instance.DONE THEN #SQCR := #STEP_85; END_IF;
END_REGION

REGION Network 26: STEP 85 TRCV
   RUNG wire#powerrail
      Contact( "AUTOMAT" )
      { S7_Templates := "SrcType := Int" } EQ_Contact(in1 := #STEP_85, in2 := #SQCR)
      wire#w1
      Contact( #TRCV_Instance.NDR )
      wire#w2
      Move(in := #STEP_90, out1 => #SQCR)
   END_RUNG
   RUNG wire#w1
      Contact( "SMAZ_ME_1" )
   END_RUNG wire#w2
   // the same network as SCL:
   IF "AUTOMAT" AND (#STEP_85 = #SQCR) AND (#TRCV_Instance.NDR OR "SMAZ_ME_1") THEN
       #SQCR := #STEP_90;
   END_IF;
END_REGION

REGION Network 27: STEP 90 DISCONNECT
   RUNG wire#powerrail
      Contact( "AUTOMAT" )
      { S7_Templates := "SrcType := Int" } EQ_Contact(in1 := #STEP_90, in2 := #SQCR)
      Contact( #TDISCON_Instance.DONE )
      Move(in := #STEP_93, out1 => #SQCR)
   END_RUNG
   // the same network as SCL:
   IF "AUTOMAT" AND (#STEP_90 = #SQCR) AND #TDISCON_Instance.DONE THEN #SQCR := #STEP_93; END_IF;
END_REGION

REGION Network 28: STEP 93 PAUZA NA VZAPAMATOVÁNÍ
   #"TIMER".TIMER_3.TON(IN := "AUTOMAT" AND (#STEP_93 = #SQCR), PT := t#500ms);
   IF #"TIMER".TIMER_3.Q THEN #SQCR := #STEP_130; END_IF;
END_REGION

REGION Network 29 (SCL): JEDEN RAMEC
   IF #Tisk.jeden_ramec AND #SQCR = #STEP_130 THEN
       #SQCR := #STEP_95;
   END_IF;
END_REGION

REGION Network 30: STEP 95 CONNECT
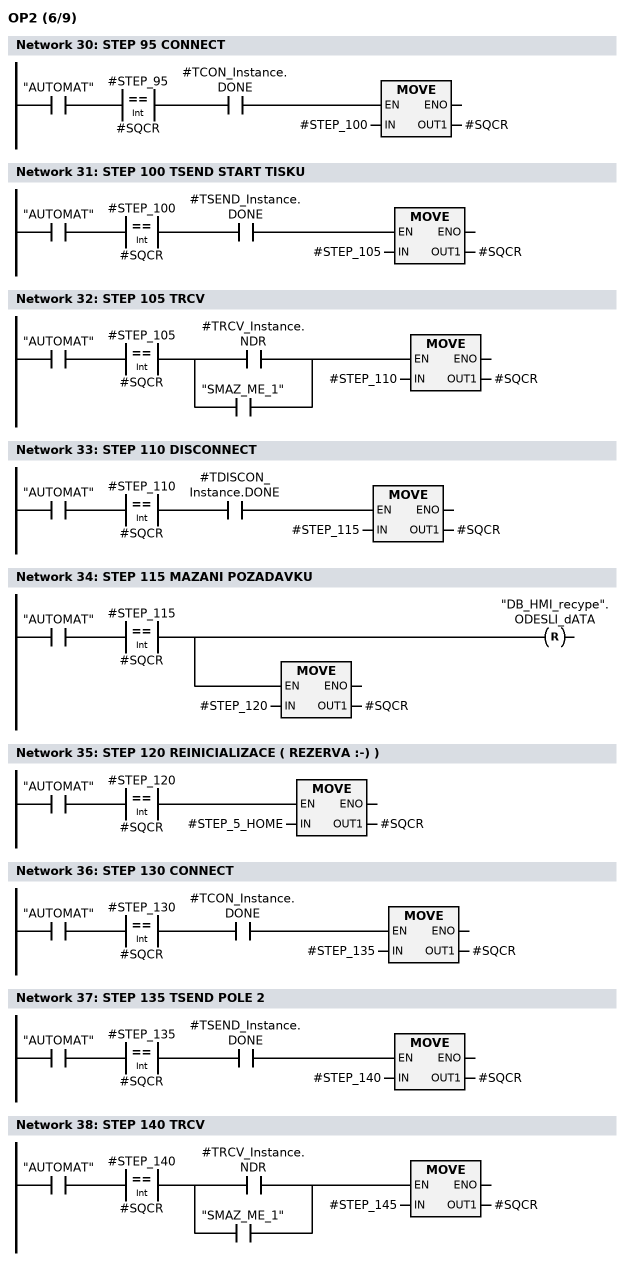
   RUNG wire#powerrail
      Contact( "AUTOMAT" )
      { S7_Templates := "SrcType := Int" } EQ_Contact(in1 := #STEP_95, in2 := #SQCR)
      Contact( #TCON_Instance.DONE )
      Move(in := #STEP_100, out1 => #SQCR)
   END_RUNG
   // the same network as SCL:
   IF "AUTOMAT" AND (#STEP_95 = #SQCR) AND #TCON_Instance.DONE THEN #SQCR := #STEP_100; END_IF;
END_REGION

REGION Network 31: STEP 100 TSEND START TISKU
   RUNG wire#powerrail
      Contact( "AUTOMAT" )
      { S7_Templates := "SrcType := Int" } EQ_Contact(in1 := #STEP_100, in2 := #SQCR)
      Contact( #TSEND_Instance.DONE )
      Move(in := #STEP_105, out1 => #SQCR)
   END_RUNG
   // the same network as SCL:
   IF "AUTOMAT" AND (#STEP_100 = #SQCR) AND #TSEND_Instance.DONE THEN #SQCR := #STEP_105; END_IF;
END_REGION

REGION Network 32: STEP 105 TRCV
   RUNG wire#powerrail
      Contact( "AUTOMAT" )
      { S7_Templates := "SrcType := Int" } EQ_Contact(in1 := #STEP_105, in2 := #SQCR)
      wire#w1
      Contact( #TRCV_Instance.NDR )
      wire#w2
      Move(in := #STEP_110, out1 => #SQCR)
   END_RUNG
   RUNG wire#w1
      Contact( "SMAZ_ME_1" )
   END_RUNG wire#w2
   // the same network as SCL:
   IF "AUTOMAT" AND (#STEP_105 = #SQCR) AND (#TRCV_Instance.NDR OR "SMAZ_ME_1") THEN
       #SQCR := #STEP_110;
   END_IF;
END_REGION

REGION Network 33: STEP 110 DISCONNECT
   RUNG wire#powerrail
      Contact( "AUTOMAT" )
      { S7_Templates := "SrcType := Int" } EQ_Contact(in1 := #STEP_110, in2 := #SQCR)
      Contact( #TDISCON_Instance.DONE )
      Move(in := #STEP_115, out1 => #SQCR)
   END_RUNG
   // the same network as SCL:
   IF "AUTOMAT" AND (#STEP_110 = #SQCR) AND #TDISCON_Instance.DONE THEN #SQCR := #STEP_115; END_IF;
END_REGION

REGION Network 34: STEP 115 MAZANI POZADAVKU
   RUNG wire#powerrail
      Contact( "AUTOMAT" )
      { S7_Templates := "SrcType := Int" } EQ_Contact(in1 := #STEP_115, in2 := #SQCR)
      wire#w1
      R_Coil( "DB_HMI_recype".ODESLI_dATA )
   END_RUNG
   RUNG wire#w1
      Move(in := #STEP_120, out1 => #SQCR)
   END_RUNG
   // the same network as SCL:
   IF "AUTOMAT" AND (#STEP_115 = #SQCR) THEN
       "DB_HMI_recype".ODESLI_dATA := FALSE;
       #SQCR := #STEP_120;
   END_IF;
END_REGION

REGION Network 35: STEP 120 REINICIALIZACE ( REZERVA :-) )
   RUNG wire#powerrail
      Contact( "AUTOMAT" )
      { S7_Templates := "SrcType := Int" } EQ_Contact(in1 := #STEP_120, in2 := #SQCR)
      Move(in := #STEP_5_HOME, out1 => #SQCR)
   END_RUNG
   // the same network as SCL:
   IF "AUTOMAT" AND (#STEP_120 = #SQCR) THEN #SQCR := #STEP_5_HOME; END_IF;
END_REGION

REGION Network 36: STEP 130 CONNECT
   RUNG wire#powerrail
      Contact( "AUTOMAT" )
      { S7_Templates := "SrcType := Int" } EQ_Contact(in1 := #STEP_130, in2 := #SQCR)
      Contact( #TCON_Instance.DONE )
      Move(in := #STEP_135, out1 => #SQCR)
   END_RUNG
   // the same network as SCL:
   IF "AUTOMAT" AND (#STEP_130 = #SQCR) AND #TCON_Instance.DONE THEN #SQCR := #STEP_135; END_IF;
END_REGION

REGION Network 37: STEP 135 TSEND POLE 2
   RUNG wire#powerrail
      Contact( "AUTOMAT" )
      { S7_Templates := "SrcType := Int" } EQ_Contact(in1 := #STEP_135, in2 := #SQCR)
      Contact( #TSEND_Instance.DONE )
      Move(in := #STEP_140, out1 => #SQCR)
   END_RUNG
   // the same network as SCL:
   IF "AUTOMAT" AND (#STEP_135 = #SQCR) AND #TSEND_Instance.DONE THEN #SQCR := #STEP_140; END_IF;
END_REGION

REGION Network 38: STEP 140 TRCV
   RUNG wire#powerrail
      Contact( "AUTOMAT" )
      { S7_Templates := "SrcType := Int" } EQ_Contact(in1 := #STEP_140, in2 := #SQCR)
      wire#w1
      Contact( #TRCV_Instance.NDR )
      wire#w2
      Move(in := #STEP_145, out1 => #SQCR)
   END_RUNG
   RUNG wire#w1
      Contact( "SMAZ_ME_1" )
   END_RUNG wire#w2
   // the same network as SCL:
   IF "AUTOMAT" AND (#STEP_140 = #SQCR) AND (#TRCV_Instance.NDR OR "SMAZ_ME_1") THEN
       #SQCR := #STEP_145;
   END_IF;
END_REGION

REGION Network 39: STEP 145 DISCONNECT
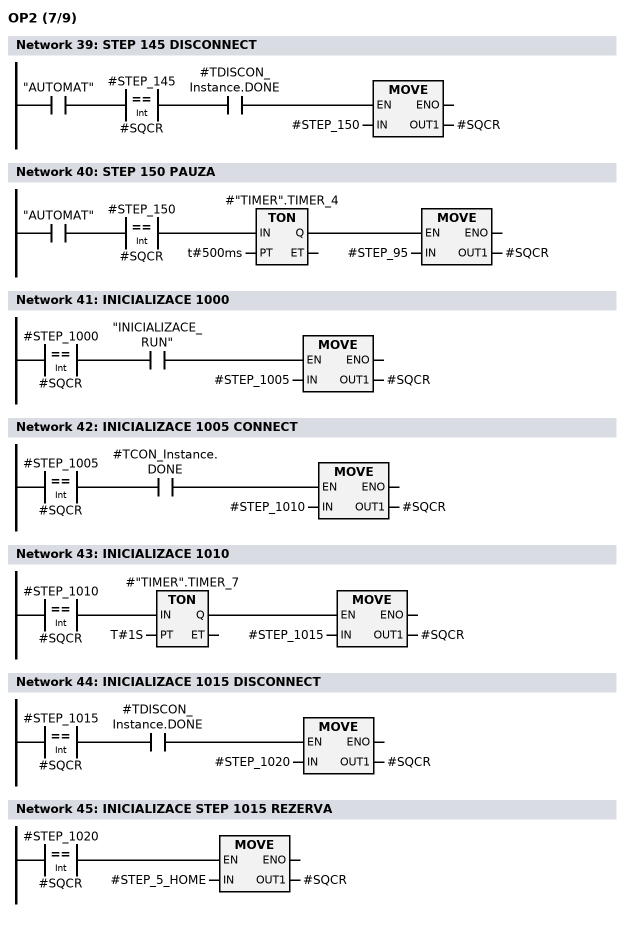
   RUNG wire#powerrail
      Contact( "AUTOMAT" )
      { S7_Templates := "SrcType := Int" } EQ_Contact(in1 := #STEP_145, in2 := #SQCR)
      Contact( #TDISCON_Instance.DONE )
      Move(in := #STEP_150, out1 => #SQCR)
   END_RUNG
   // the same network as SCL:
   IF "AUTOMAT" AND (#STEP_145 = #SQCR) AND #TDISCON_Instance.DONE THEN #SQCR := #STEP_150; END_IF;
END_REGION

REGION Network 40: STEP 150 PAUZA
   #"TIMER".TIMER_4.TON(IN := "AUTOMAT" AND (#STEP_150 = #SQCR), PT := t#500ms);
   IF #"TIMER".TIMER_4.Q THEN #SQCR := #STEP_95; END_IF;
END_REGION

REGION Network 41: INICIALIZACE 1000
   RUNG wire#powerrail
      { S7_Templates := "SrcType := Int" } EQ_Contact(in1 := #STEP_1000, in2 := #SQCR)
      Contact( "INICIALIZACE_RUN" )
      Move(in := #STEP_1005, out1 => #SQCR)
   END_RUNG
   // the same network as SCL:
   IF (#STEP_1000 = #SQCR) AND "INICIALIZACE_RUN" THEN #SQCR := #STEP_1005; END_IF;
END_REGION

REGION Network 42: INICIALIZACE 1005 CONNECT
   RUNG wire#powerrail
      { S7_Templates := "SrcType := Int" } EQ_Contact(in1 := #STEP_1005, in2 := #SQCR)
      Contact( #TCON_Instance.DONE )
      Move(in := #STEP_1010, out1 => #SQCR)
   END_RUNG
   // the same network as SCL:
   IF (#STEP_1005 = #SQCR) AND #TCON_Instance.DONE THEN #SQCR := #STEP_1010; END_IF;
END_REGION

REGION Network 43: INICIALIZACE 1010
   #"TIMER".TIMER_7.TON(IN := #STEP_1010 = #SQCR, PT := T#1S);
   IF #"TIMER".TIMER_7.Q THEN #SQCR := #STEP_1015; END_IF;
END_REGION

REGION Network 44: INICIALIZACE 1015 DISCONNECT
   RUNG wire#powerrail
      { S7_Templates := "SrcType := Int" } EQ_Contact(in1 := #STEP_1015, in2 := #SQCR)
      Contact( #TDISCON_Instance.DONE )
      Move(in := #STEP_1020, out1 => #SQCR)
   END_RUNG
   // the same network as SCL:
   IF (#STEP_1015 = #SQCR) AND #TDISCON_Instance.DONE THEN #SQCR := #STEP_1020; END_IF;
END_REGION

REGION Network 45: INICIALIZACE STEP 1015 REZERVA
   RUNG wire#powerrail
      { S7_Templates := "SrcType := Int" } EQ_Contact(in1 := #STEP_1020, in2 := #SQCR)
      Move(in := #STEP_5_HOME, out1 => #SQCR)
   END_RUNG
   // the same network as SCL:
   IF #STEP_1020 = #SQCR THEN #SQCR := #STEP_5_HOME; END_IF;
END_REGION

REGION Network 46: automat control tiskarna / automat control door
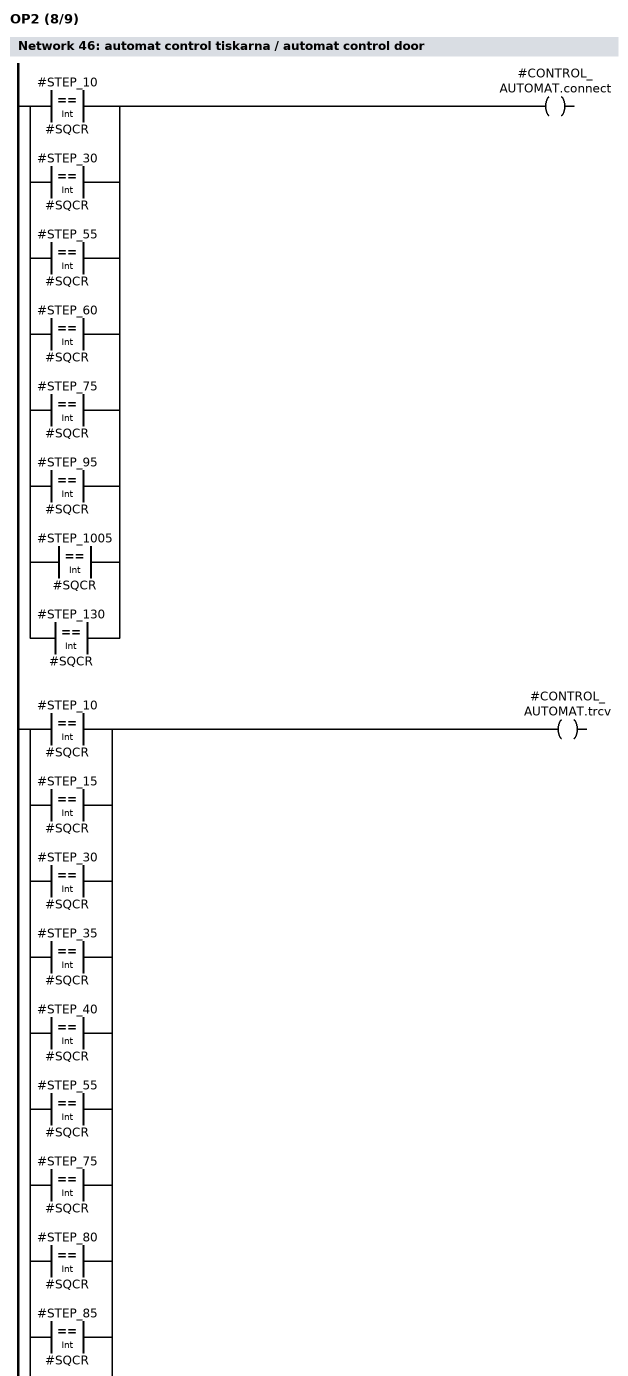
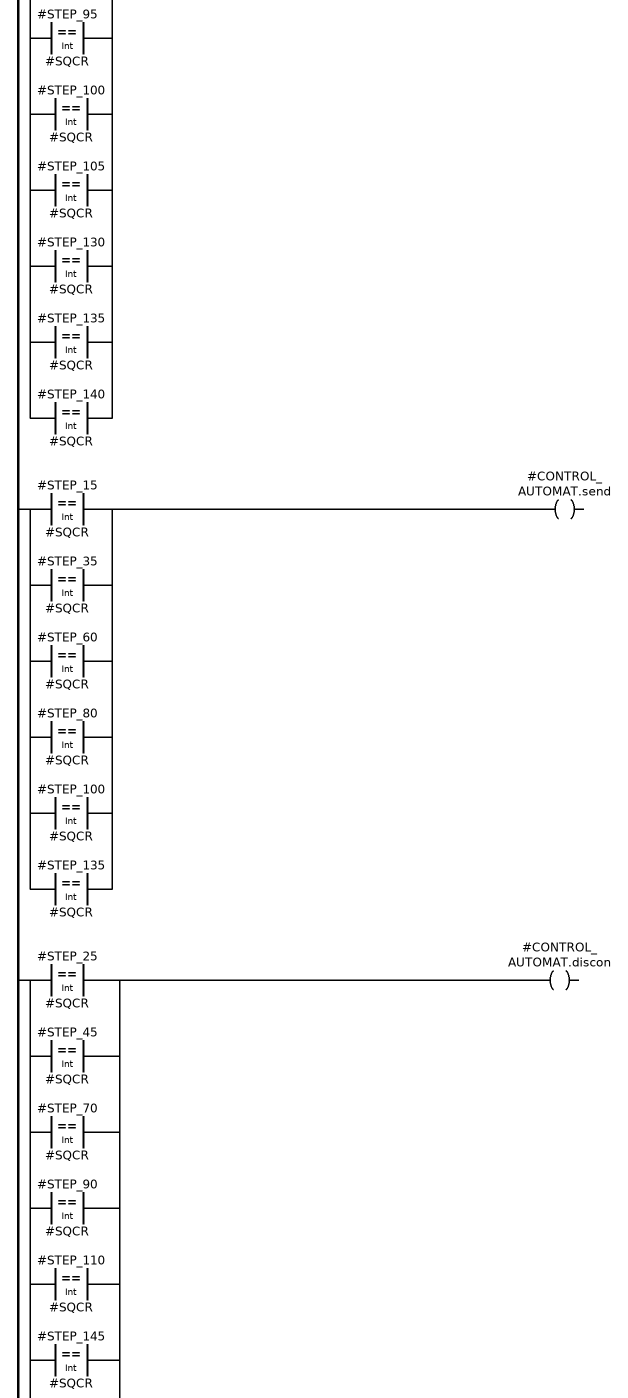
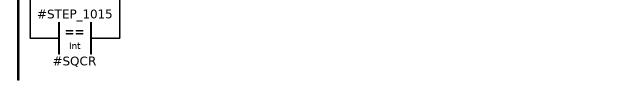
   RUNG wire#powerrail
      { S7_Templates := "SrcType := Int" } EQ_Contact(in1 := #STEP_10, in2 := #SQCR)
      wire#w1
      Coil( #CONTROL_AUTOMAT.connect )
   END_RUNG
   RUNG wire#powerrail
      { S7_Templates := "SrcType := Int" } EQ_Contact(in1 := #STEP_30, in2 := #SQCR)
   END_RUNG wire#w1
   RUNG wire#powerrail
      { S7_Templates := "SrcType := Int" } EQ_Contact(in1 := #STEP_55, in2 := #SQCR)
   END_RUNG wire#w1
   RUNG wire#powerrail
      { S7_Templates := "SrcType := Int" } EQ_Contact(in1 := #STEP_60, in2 := #SQCR)
   END_RUNG wire#w1
   RUNG wire#powerrail
      { S7_Templates := "SrcType := Int" } EQ_Contact(in1 := #STEP_75, in2 := #SQCR)
   END_RUNG wire#w1
   RUNG wire#powerrail
      { S7_Templates := "SrcType := Int" } EQ_Contact(in1 := #STEP_95, in2 := #SQCR)
   END_RUNG wire#w1
   RUNG wire#powerrail
      { S7_Templates := "SrcType := Int" } EQ_Contact(in1 := #STEP_1005, in2 := #SQCR)
   END_RUNG wire#w1
   RUNG wire#powerrail
      { S7_Templates := "SrcType := Int" } EQ_Contact(in1 := #STEP_130, in2 := #SQCR)
   END_RUNG wire#w1
   RUNG wire#powerrail
      { S7_Templates := "SrcType := Int" } EQ_Contact(in1 := #STEP_10, in2 := #SQCR)
      wire#w2
      Coil( #CONTROL_AUTOMAT.trcv )
   END_RUNG
   RUNG wire#powerrail
      { S7_Templates := "SrcType := Int" } EQ_Contact(in1 := #STEP_15, in2 := #SQCR)
   END_RUNG wire#w2
   RUNG wire#powerrail
      { S7_Templates := "SrcType := Int" } EQ_Contact(in1 := #STEP_30, in2 := #SQCR)
   END_RUNG wire#w2
   RUNG wire#powerrail
      { S7_Templates := "SrcType := Int" } EQ_Contact(in1 := #STEP_35, in2 := #SQCR)
   END_RUNG wire#w2
   RUNG wire#powerrail
      { S7_Templates := "SrcType := Int" } EQ_Contact(in1 := #STEP_40, in2 := #SQCR)
   END_RUNG wire#w2
   RUNG wire#powerrail
      { S7_Templates := "SrcType := Int" } EQ_Contact(in1 := #STEP_55, in2 := #SQCR)
   END_RUNG wire#w2
   RUNG wire#powerrail
      { S7_Templates := "SrcType := Int" } EQ_Contact(in1 := #STEP_75, in2 := #SQCR)
   END_RUNG wire#w2
   RUNG wire#powerrail
      { S7_Templates := "SrcType := Int" } EQ_Contact(in1 := #STEP_80, in2 := #SQCR)
   END_RUNG wire#w2
   RUNG wire#powerrail
      { S7_Templates := "SrcType := Int" } EQ_Contact(in1 := #STEP_85, in2 := #SQCR)
   END_RUNG wire#w2
   RUNG wire#powerrail
      { S7_Templates := "SrcType := Int" } EQ_Contact(in1 := #STEP_95, in2 := #SQCR)
   END_RUNG wire#w2
   RUNG wire#powerrail
      { S7_Templates := "SrcType := Int" } EQ_Contact(in1 := #STEP_100, in2 := #SQCR)
   END_RUNG wire#w2
   RUNG wire#powerrail
      { S7_Templates := "SrcType := Int" } EQ_Contact(in1 := #STEP_105, in2 := #SQCR)
   END_RUNG wire#w2
   RUNG wire#powerrail
      { S7_Templates := "SrcType := Int" } EQ_Contact(in1 := #STEP_130, in2 := #SQCR)
   END_RUNG wire#w2
   RUNG wire#powerrail
      { S7_Templates := "SrcType := Int" } EQ_Contact(in1 := #STEP_135, in2 := #SQCR)
   END_RUNG wire#w2
   RUNG wire#powerrail
      { S7_Templates := "SrcType := Int" } EQ_Contact(in1 := #STEP_140, in2 := #SQCR)
   END_RUNG wire#w2
   RUNG wire#powerrail
      { S7_Templates := "SrcType := Int" } EQ_Contact(in1 := #STEP_15, in2 := #SQCR)
      wire#w3
      Coil( #CONTROL_AUTOMAT.send )
   END_RUNG
   RUNG wire#powerrail
      { S7_Templates := "SrcType := Int" } EQ_Contact(in1 := #STEP_35, in2 := #SQCR)
   END_RUNG wire#w3
   RUNG wire#powerrail
      { S7_Templates := "SrcType := Int" } EQ_Contact(in1 := #STEP_60, in2 := #SQCR)
   END_RUNG wire#w3
   RUNG wire#powerrail
      { S7_Templates := "SrcType := Int" } EQ_Contact(in1 := #STEP_80, in2 := #SQCR)
   END_RUNG wire#w3
   RUNG wire#powerrail
      { S7_Templates := "SrcType := Int" } EQ_Contact(in1 := #STEP_100, in2 := #SQCR)
   END_RUNG wire#w3
   RUNG wire#powerrail
      { S7_Templates := "SrcType := Int" } EQ_Contact(in1 := #STEP_135, in2 := #SQCR)
   END_RUNG wire#w3
   RUNG wire#powerrail
      { S7_Templates := "SrcType := Int" } EQ_Contact(in1 := #STEP_25, in2 := #SQCR)
      wire#w4
      Coil( #CONTROL_AUTOMAT.discon )
   END_RUNG
   RUNG wire#powerrail
      { S7_Templates := "SrcType := Int" } EQ_Contact(in1 := #STEP_45, in2 := #SQCR)
   END_RUNG wire#w4
   RUNG wire#powerrail
      { S7_Templates := "SrcType := Int" } EQ_Contact(in1 := #STEP_70, in2 := #SQCR)
   END_RUNG wire#w4
   RUNG wire#powerrail
      { S7_Templates := "SrcType := Int" } EQ_Contact(in1 := #STEP_90, in2 := #SQCR)
   END_RUNG wire#w4
   RUNG wire#powerrail
      { S7_Templates := "SrcType := Int" } EQ_Contact(in1 := #STEP_110, in2 := #SQCR)
   END_RUNG wire#w4
   RUNG wire#powerrail
      { S7_Templates := "SrcType := Int" } EQ_Contact(in1 := #STEP_145, in2 := #SQCR)
   END_RUNG wire#w4
   RUNG wire#powerrail
      { S7_Templates := "SrcType := Int" } EQ_Contact(in1 := #STEP_1015, in2 := #SQCR)
   END_RUNG wire#w4
   // the same network as SCL:
   #CONTROL_AUTOMAT.connect := (#STEP_10 = #SQCR) OR (#STEP_30 = #SQCR) OR (#STEP_55 = #SQCR) OR (#STEP_60 = #SQCR) OR (#STEP_75 = #SQCR) OR (#STEP_95 = #SQCR) OR (#STEP_1005 = #SQCR) OR (#STEP_130 = #SQCR);
   #CONTROL_AUTOMAT.trcv := (#STEP_10 = #SQCR) OR (#STEP_15 = #SQCR) OR (#STEP_30 = #SQCR) OR (#STEP_35 = #SQCR) OR (#STEP_40 = #SQCR) OR (#STEP_55 = #SQCR) OR (#STEP_75 = #SQCR) OR (#STEP_80 = #SQCR) OR (#STEP_85 = #SQCR) OR (#STEP_95 = #SQCR) OR (#STEP_100 = #SQCR) OR (#STEP_105 = #SQCR) OR (#STEP_130 = #SQCR) OR (#STEP_135 = #SQCR) OR (#STEP_140 = #SQCR);
   #CONTROL_AUTOMAT.send := (#STEP_15 = #SQCR) OR (#STEP_35 = #SQCR) OR (#STEP_60 = #SQCR) OR (#STEP_80 = #SQCR) OR (#STEP_100 = #SQCR) OR (#STEP_135 = #SQCR);
   #CONTROL_AUTOMAT.discon := (#STEP_25 = #SQCR) OR (#STEP_45 = #SQCR) OR (#STEP_70 = #SQCR) OR (#STEP_90 = #SQCR) OR (#STEP_110 = #SQCR) OR (#STEP_145 = #SQCR) OR (#STEP_1015 = #SQCR);
END_REGION

REGION Network 47: EXTERNAL_TRIGER
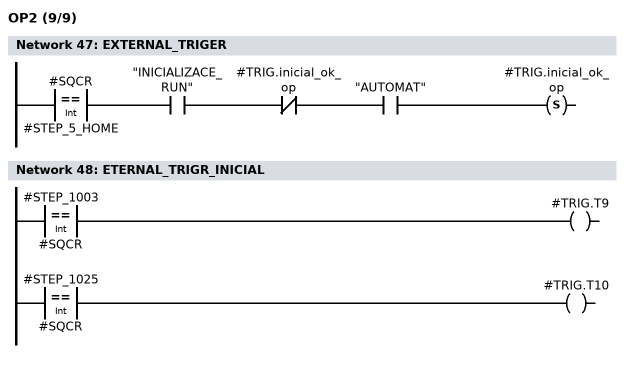
   RUNG wire#powerrail
      { S7_Templates := "SrcType := Int" } EQ_Contact(in1 := #SQCR, in2 := #STEP_5_HOME)
      Contact( "INICIALIZACE_RUN" )
      I_Contact( #TRIG.inicial_ok_op )
      Contact( "AUTOMAT" )
      S_Coil( #TRIG.inicial_ok_op )
   END_RUNG
   // the same network as SCL:
   IF (#SQCR = #STEP_5_HOME) AND "INICIALIZACE_RUN" AND NOT #TRIG.inicial_ok_op AND "AUTOMAT" THEN
       #TRIG.inicial_ok_op := TRUE;
   END_IF;
END_REGION

REGION Network 48: ETERNAL_TRIGR_INICIAL
   RUNG wire#powerrail
      { S7_Templates := "SrcType := Int" } EQ_Contact(in1 := #STEP_1003, in2 := #SQCR)
      Coil( #TRIG.T9 )
   END_RUNG
   RUNG wire#powerrail
      { S7_Templates := "SrcType := Int" } EQ_Contact(in1 := #STEP_1025, in2 := #SQCR)
      Coil( #TRIG.T10 )
   END_RUNG
   // the same network as SCL:
   #TRIG.T9 := #STEP_1003 = #SQCR;
   #TRIG.T10 := #STEP_1025 = #SQCR;
END_REGION

REGION Network 49: hmi
END_REGION
END_FUNCTION_BLOCK

// folder: OPERACE/MANUAL CONTROL

FUNCTION_BLOCK "FB_CamManual"   // FB1, SCL
{ S7_Optimized_Access := 'TRUE' }
VERSION : 0.1
   VAR_INPUT
      xManEtiketa : Bool;   // ruční test etiketa
      xManFolie : Bool;   // ruční test folie
      tLightDelay : Time := T#100ms;   // náběh světel
      tTrigPulse : Time := T#50ms;   // d0lka triggeru
   END_VAR
   VAR
      tonEt : TON_TIME;
      tpEt : TP_TIME;
      tonFo : TON_TIME;
      tpFo : TP_TIME;
   END_VAR
BEGIN
   // ---------- ETIKETA ----------
   #tonEt(IN := #xManEtiketa,
          PT := #tLightDelay);
   #tpEt(IN := #tonEt.Q,
         PT := #tTrigPulse);

   IF #xManEtiketa THEN
       "-KA1" := TRUE;
       "-KA2" := TRUE;
   END_IF;
   IF #tpEt.Q THEN
       "COG_ETIKETA_COG_ETIKETA_is3800-Trigger" := TRUE;
   END_IF;

   // ---------- FÓLIE ----------
   #tonFo(IN := #xManFolie,
          PT := #tLightDelay);
   #tpFo(IN := #tonFo.Q,
         PT := #tTrigPulse);

   IF #xManFolie THEN
       "-KA3" := TRUE;
       "-KA4" := TRUE;
       "-KA5" := TRUE;
   END_IF;
   IF #tpFo.Q THEN
       "COG_FOLIE_L_is3800-Trigger" := TRUE;
       "COG_FOLIE_P_is3800-Trigger" := TRUE;
   END_IF;
END_FUNCTION_BLOCK

FUNCTION "FC_PocetChyb" : Int   // FC2, SCL
{ S7_Optimized_Access := 'TRUE' }
VERSION : 0.1
   VAR_INPUT
      "A" : String;
      "B" : String;
   END_VAR
   VAR_TEMP
      la : Int;
      lb : Int;
      i : Int;
      j : Int;
      v : Int;
      prev : Array[0..40] of Int;
      cur : Array[0..40] of Int;
   END_VAR
BEGIN
   // Pocet chyb mezi texty A a B (kolik znaku zamenit / vlozit / smazat).
   // 0 = texty jsou shodne. Porovnava se max. 40 znaku kvuli dobe cyklu.
   #la := MIN(IN1 := LEN(#A), IN2 := 40);
   #lb := MIN(IN1 := LEN(#B), IN2 := 40);

   FOR #j := 0 TO #lb DO
       #prev[#j] := #j;
   END_FOR;

   FOR #i := 1 TO #la DO
       #cur[0] := #i;
       FOR #j := 1 TO #lb DO
           #v := #prev[#j - 1];                // shoda / zamena znaku
           IF #A[#i] <> #B[#j] THEN
               #v := #v + 1;
           END_IF;
           IF #prev[#j] + 1 < #v THEN          // znak navic
               #v := #prev[#j] + 1;
           END_IF;
           IF #cur[#j - 1] + 1 < #v THEN       // chybejici znak
               #v := #cur[#j - 1] + 1;
           END_IF;
           #cur[#j] := #v;
       END_FOR;
       FOR #j := 0 TO #lb DO
           #prev[#j] := #cur[#j];
       END_FOR;
   END_FOR;

   #FC_PocetChyb := #prev[#lb];
END_FUNCTION

// folder: STANDARD/ALARM

FUNCTION "alarmy" : Void   // FC100, LAD
{ S7_Optimized_Access := 'TRUE' }
VERSION : 0.1
   VAR_OUTPUT
      fc_alarm_global : Bool;
      fc_wrong_global : Bool;
      fc_op_1_alrm : Bool;
      fc_op_1_wrong : Bool;
      fc_op_2_alrm : Bool;
      fc_op_2_wrong : Bool;
      fc_op_3_alrm : Bool;
      fc_op_3_wrong : Bool;
   END_VAR
   VAR_TEMP
      OP_1_E : Bool;
      OP_2_E : Bool;
      OP_3_E : Bool;
      OP_4_E : Bool;
      OP_5_E : Bool;
      OP_1_W : Bool;
      OP_2_W : Bool;
      OP_3_W : Bool;
      OP_4_W : Bool;
      OP_5_W : Bool;
   END_VAR
   VAR CONSTANT
      TIME_ERROR_BOR : Time := T#4S;
   END_VAR
BEGIN

REGION Network 1: op_1 alarmy proces
END_REGION

REGION Network 2: op_1_warning_proces
END_REGION

REGION Network 3: OP_1_ALARM
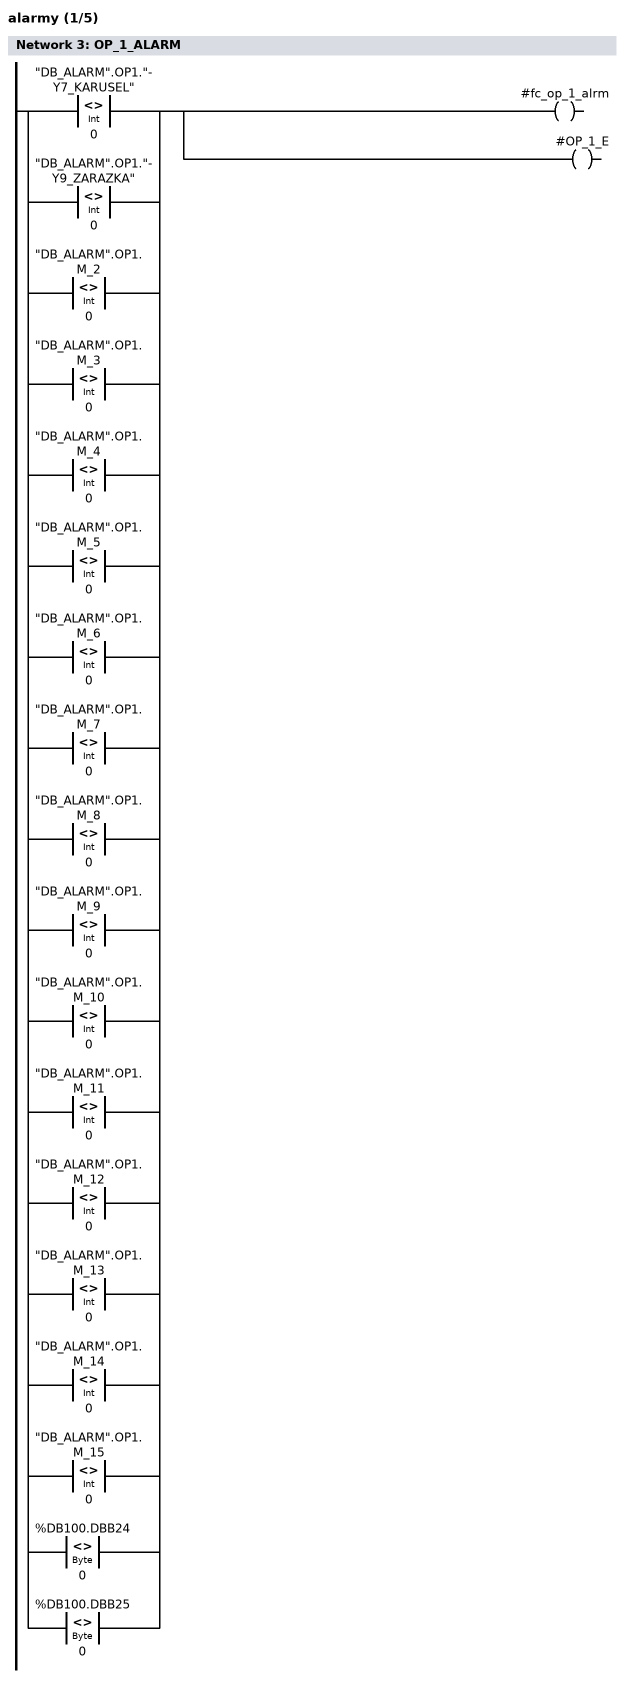
   RUNG wire#powerrail
      { S7_Templates := "SrcType := Int" } NE_Contact(in1 := "DB_ALARM".OP1."-Y7_KARUSEL", in2 := 0)
      wire#w1
      Coil( #fc_op_1_alrm )
   END_RUNG
   RUNG wire#powerrail
      { S7_Templates := "SrcType := Int" } NE_Contact(in1 := "DB_ALARM".OP1."-Y9_ZARAZKA", in2 := 0)
   END_RUNG wire#w1
   RUNG wire#powerrail
      { S7_Templates := "SrcType := Int" } NE_Contact(in1 := "DB_ALARM".OP1.M_2, in2 := 0)
   END_RUNG wire#w1
   RUNG wire#powerrail
      { S7_Templates := "SrcType := Int" } NE_Contact(in1 := "DB_ALARM".OP1.M_3, in2 := 0)
   END_RUNG wire#w1
   RUNG wire#powerrail
      { S7_Templates := "SrcType := Int" } NE_Contact(in1 := "DB_ALARM".OP1.M_4, in2 := 0)
   END_RUNG wire#w1
   RUNG wire#powerrail
      { S7_Templates := "SrcType := Int" } NE_Contact(in1 := "DB_ALARM".OP1.M_5, in2 := 0)
   END_RUNG wire#w1
   RUNG wire#powerrail
      { S7_Templates := "SrcType := Int" } NE_Contact(in1 := "DB_ALARM".OP1.M_6, in2 := 0)
   END_RUNG wire#w1
   RUNG wire#powerrail
      { S7_Templates := "SrcType := Int" } NE_Contact(in1 := "DB_ALARM".OP1.M_7, in2 := 0)
   END_RUNG wire#w1
   RUNG wire#powerrail
      { S7_Templates := "SrcType := Int" } NE_Contact(in1 := "DB_ALARM".OP1.M_8, in2 := 0)
   END_RUNG wire#w1
   RUNG wire#powerrail
      { S7_Templates := "SrcType := Int" } NE_Contact(in1 := "DB_ALARM".OP1.M_9, in2 := 0)
   END_RUNG wire#w1
   RUNG wire#powerrail
      { S7_Templates := "SrcType := Int" } NE_Contact(in1 := "DB_ALARM".OP1.M_10, in2 := 0)
   END_RUNG wire#w1
   RUNG wire#powerrail
      { S7_Templates := "SrcType := Int" } NE_Contact(in1 := "DB_ALARM".OP1.M_11, in2 := 0)
   END_RUNG wire#w1
   RUNG wire#powerrail
      { S7_Templates := "SrcType := Int" } NE_Contact(in1 := "DB_ALARM".OP1.M_12, in2 := 0)
   END_RUNG wire#w1
   RUNG wire#powerrail
      { S7_Templates := "SrcType := Int" } NE_Contact(in1 := "DB_ALARM".OP1.M_13, in2 := 0)
   END_RUNG wire#w1
   RUNG wire#powerrail
      { S7_Templates := "SrcType := Int" } NE_Contact(in1 := "DB_ALARM".OP1.M_14, in2 := 0)
   END_RUNG wire#w1
   RUNG wire#powerrail
      { S7_Templates := "SrcType := Int" } NE_Contact(in1 := "DB_ALARM".OP1.M_15, in2 := 0)
   END_RUNG wire#w1
   RUNG wire#powerrail
      { S7_Templates := "SrcType := Byte" } NE_Contact(in1 := %DB100.DBB24, in2 := 0)
   END_RUNG wire#w1
   RUNG wire#powerrail
      { S7_Templates := "SrcType := Byte" } NE_Contact(in1 := %DB100.DBB25, in2 := 0)
   END_RUNG wire#w1
   RUNG wire#w1
      Coil( #OP_1_E )
   END_RUNG
   // the same network as SCL:
   #fc_op_1_alrm := ("DB_ALARM".OP1."-Y7_KARUSEL" <> 0) OR ("DB_ALARM".OP1."-Y9_ZARAZKA" <> 0) OR ("DB_ALARM".OP1.M_2 <> 0) OR ("DB_ALARM".OP1.M_3 <> 0) OR ("DB_ALARM".OP1.M_4 <> 0) OR ("DB_ALARM".OP1.M_5 <> 0) OR ("DB_ALARM".OP1.M_6 <> 0) OR ("DB_ALARM".OP1.M_7 <> 0) OR ("DB_ALARM".OP1.M_8 <> 0) OR ("DB_ALARM".OP1.M_9 <> 0) OR ("DB_ALARM".OP1.M_10 <> 0) OR ("DB_ALARM".OP1.M_11 <> 0) OR ("DB_ALARM".OP1.M_12 <> 0) OR ("DB_ALARM".OP1.M_13 <> 0) OR ("DB_ALARM".OP1.M_14 <> 0) OR ("DB_ALARM".OP1.M_15 <> 0) OR (%DB100.DBB24 <> 0) OR (%DB100.DBB25 <> 0);
   #OP_1_E := #fc_op_1_alrm;
END_REGION

REGION Network 4: OP_2_ALARM
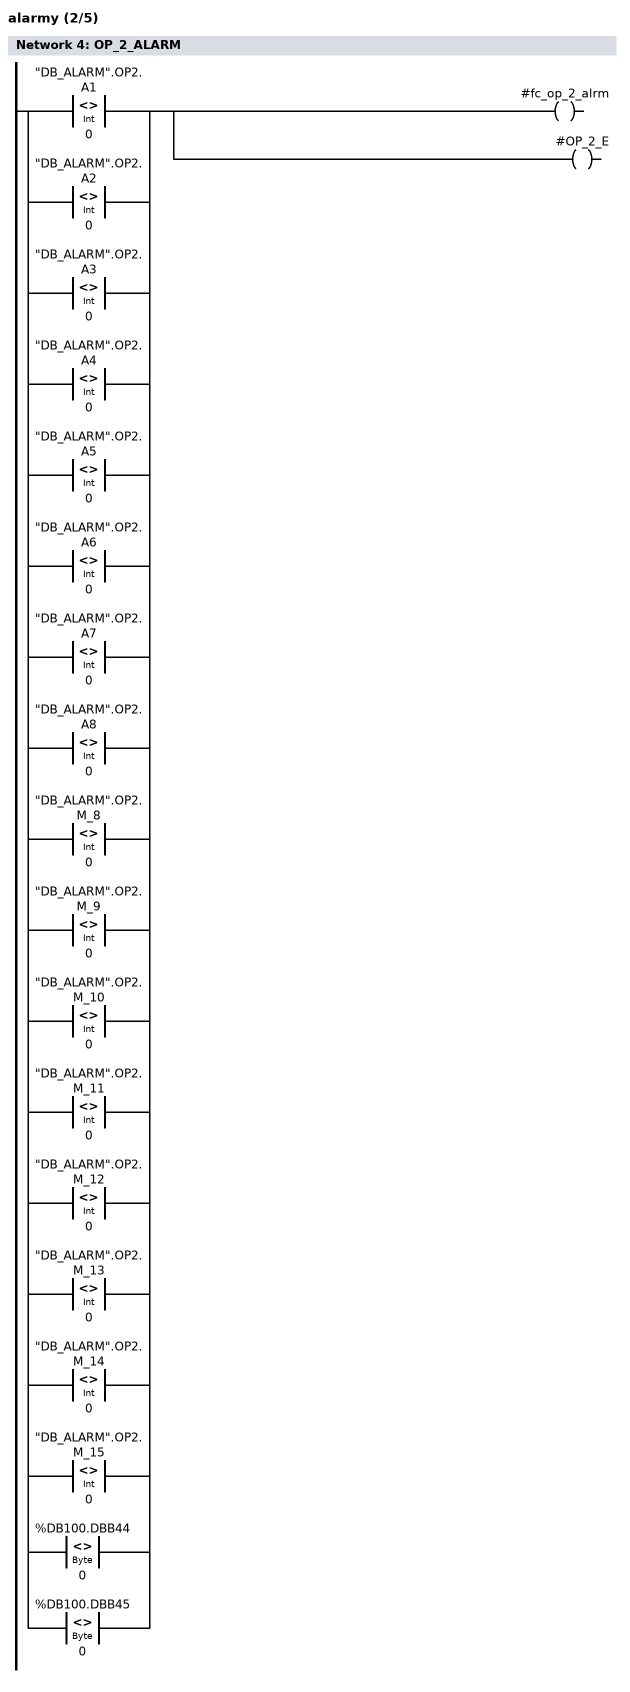
   RUNG wire#powerrail
      { S7_Templates := "SrcType := Int" } NE_Contact(in1 := "DB_ALARM".OP2.A1, in2 := 0)
      wire#w1
      Coil( #fc_op_2_alrm )
   END_RUNG
   RUNG wire#powerrail
      { S7_Templates := "SrcType := Int" } NE_Contact(in1 := "DB_ALARM".OP2.A2, in2 := 0)
   END_RUNG wire#w1
   RUNG wire#powerrail
      { S7_Templates := "SrcType := Int" } NE_Contact(in1 := "DB_ALARM".OP2.A3, in2 := 0)
   END_RUNG wire#w1
   RUNG wire#powerrail
      { S7_Templates := "SrcType := Int" } NE_Contact(in1 := "DB_ALARM".OP2.A4, in2 := 0)
   END_RUNG wire#w1
   RUNG wire#powerrail
      { S7_Templates := "SrcType := Int" } NE_Contact(in1 := "DB_ALARM".OP2.A5, in2 := 0)
   END_RUNG wire#w1
   RUNG wire#powerrail
      { S7_Templates := "SrcType := Int" } NE_Contact(in1 := "DB_ALARM".OP2.A6, in2 := 0)
   END_RUNG wire#w1
   RUNG wire#powerrail
      { S7_Templates := "SrcType := Int" } NE_Contact(in1 := "DB_ALARM".OP2.A7, in2 := 0)
   END_RUNG wire#w1
   RUNG wire#powerrail
      { S7_Templates := "SrcType := Int" } NE_Contact(in1 := "DB_ALARM".OP2.A8, in2 := 0)
   END_RUNG wire#w1
   RUNG wire#powerrail
      { S7_Templates := "SrcType := Int" } NE_Contact(in1 := "DB_ALARM".OP2.M_8, in2 := 0)
   END_RUNG wire#w1
   RUNG wire#powerrail
      { S7_Templates := "SrcType := Int" } NE_Contact(in1 := "DB_ALARM".OP2.M_9, in2 := 0)
   END_RUNG wire#w1
   RUNG wire#powerrail
      { S7_Templates := "SrcType := Int" } NE_Contact(in1 := "DB_ALARM".OP2.M_10, in2 := 0)
   END_RUNG wire#w1
   RUNG wire#powerrail
      { S7_Templates := "SrcType := Int" } NE_Contact(in1 := "DB_ALARM".OP2.M_11, in2 := 0)
   END_RUNG wire#w1
   RUNG wire#powerrail
      { S7_Templates := "SrcType := Int" } NE_Contact(in1 := "DB_ALARM".OP2.M_12, in2 := 0)
   END_RUNG wire#w1
   RUNG wire#powerrail
      { S7_Templates := "SrcType := Int" } NE_Contact(in1 := "DB_ALARM".OP2.M_13, in2 := 0)
   END_RUNG wire#w1
   RUNG wire#powerrail
      { S7_Templates := "SrcType := Int" } NE_Contact(in1 := "DB_ALARM".OP2.M_14, in2 := 0)
   END_RUNG wire#w1
   RUNG wire#powerrail
      { S7_Templates := "SrcType := Int" } NE_Contact(in1 := "DB_ALARM".OP2.M_15, in2 := 0)
   END_RUNG wire#w1
   RUNG wire#powerrail
      { S7_Templates := "SrcType := Byte" } NE_Contact(in1 := %DB100.DBB44, in2 := 0)
   END_RUNG wire#w1
   RUNG wire#powerrail
      { S7_Templates := "SrcType := Byte" } NE_Contact(in1 := %DB100.DBB45, in2 := 0)
   END_RUNG wire#w1
   RUNG wire#w1
      Coil( #OP_2_E )
   END_RUNG
   // the same network as SCL:
   #fc_op_2_alrm := ("DB_ALARM".OP2.A1 <> 0) OR ("DB_ALARM".OP2.A2 <> 0) OR ("DB_ALARM".OP2.A3 <> 0) OR ("DB_ALARM".OP2.A4 <> 0) OR ("DB_ALARM".OP2.A5 <> 0) OR ("DB_ALARM".OP2.A6 <> 0) OR ("DB_ALARM".OP2.A7 <> 0) OR ("DB_ALARM".OP2.A8 <> 0) OR ("DB_ALARM".OP2.M_8 <> 0) OR ("DB_ALARM".OP2.M_9 <> 0) OR ("DB_ALARM".OP2.M_10 <> 0) OR ("DB_ALARM".OP2.M_11 <> 0) OR ("DB_ALARM".OP2.M_12 <> 0) OR ("DB_ALARM".OP2.M_13 <> 0) OR ("DB_ALARM".OP2.M_14 <> 0) OR ("DB_ALARM".OP2.M_15 <> 0) OR (%DB100.DBB44 <> 0) OR (%DB100.DBB45 <> 0);
   #OP_2_E := #fc_op_2_alrm;
END_REGION

REGION Network 5: OP_3_ALARM
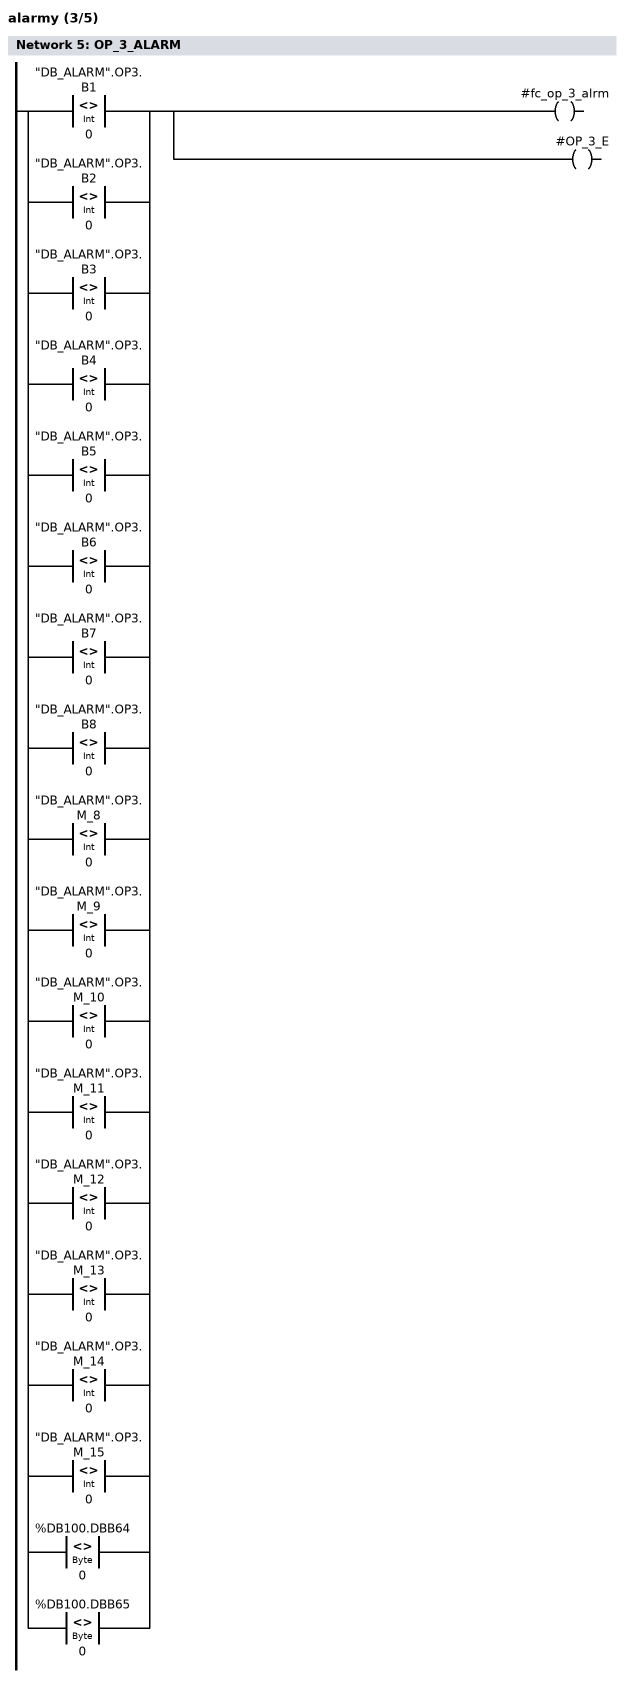
   RUNG wire#powerrail
      { S7_Templates := "SrcType := Int" } NE_Contact(in1 := "DB_ALARM".OP3.B1, in2 := 0)
      wire#w1
      Coil( #fc_op_3_alrm )
   END_RUNG
   RUNG wire#powerrail
      { S7_Templates := "SrcType := Int" } NE_Contact(in1 := "DB_ALARM".OP3.B2, in2 := 0)
   END_RUNG wire#w1
   RUNG wire#powerrail
      { S7_Templates := "SrcType := Int" } NE_Contact(in1 := "DB_ALARM".OP3.B3, in2 := 0)
   END_RUNG wire#w1
   RUNG wire#powerrail
      { S7_Templates := "SrcType := Int" } NE_Contact(in1 := "DB_ALARM".OP3.B4, in2 := 0)
   END_RUNG wire#w1
   RUNG wire#powerrail
      { S7_Templates := "SrcType := Int" } NE_Contact(in1 := "DB_ALARM".OP3.B5, in2 := 0)
   END_RUNG wire#w1
   RUNG wire#powerrail
      { S7_Templates := "SrcType := Int" } NE_Contact(in1 := "DB_ALARM".OP3.B6, in2 := 0)
   END_RUNG wire#w1
   RUNG wire#powerrail
      { S7_Templates := "SrcType := Int" } NE_Contact(in1 := "DB_ALARM".OP3.B7, in2 := 0)
   END_RUNG wire#w1
   RUNG wire#powerrail
      { S7_Templates := "SrcType := Int" } NE_Contact(in1 := "DB_ALARM".OP3.B8, in2 := 0)
   END_RUNG wire#w1
   RUNG wire#powerrail
      { S7_Templates := "SrcType := Int" } NE_Contact(in1 := "DB_ALARM".OP3.M_8, in2 := 0)
   END_RUNG wire#w1
   RUNG wire#powerrail
      { S7_Templates := "SrcType := Int" } NE_Contact(in1 := "DB_ALARM".OP3.M_9, in2 := 0)
   END_RUNG wire#w1
   RUNG wire#powerrail
      { S7_Templates := "SrcType := Int" } NE_Contact(in1 := "DB_ALARM".OP3.M_10, in2 := 0)
   END_RUNG wire#w1
   RUNG wire#powerrail
      { S7_Templates := "SrcType := Int" } NE_Contact(in1 := "DB_ALARM".OP3.M_11, in2 := 0)
   END_RUNG wire#w1
   RUNG wire#powerrail
      { S7_Templates := "SrcType := Int" } NE_Contact(in1 := "DB_ALARM".OP3.M_12, in2 := 0)
   END_RUNG wire#w1
   RUNG wire#powerrail
      { S7_Templates := "SrcType := Int" } NE_Contact(in1 := "DB_ALARM".OP3.M_13, in2 := 0)
   END_RUNG wire#w1
   RUNG wire#powerrail
      { S7_Templates := "SrcType := Int" } NE_Contact(in1 := "DB_ALARM".OP3.M_14, in2 := 0)
   END_RUNG wire#w1
   RUNG wire#powerrail
      { S7_Templates := "SrcType := Int" } NE_Contact(in1 := "DB_ALARM".OP3.M_15, in2 := 0)
   END_RUNG wire#w1
   RUNG wire#powerrail
      { S7_Templates := "SrcType := Byte" } NE_Contact(in1 := %DB100.DBB64, in2 := 0)
   END_RUNG wire#w1
   RUNG wire#powerrail
      { S7_Templates := "SrcType := Byte" } NE_Contact(in1 := %DB100.DBB65, in2 := 0)
   END_RUNG wire#w1
   RUNG wire#w1
      Coil( #OP_3_E )
   END_RUNG
   // the same network as SCL:
   #fc_op_3_alrm := ("DB_ALARM".OP3.B1 <> 0) OR ("DB_ALARM".OP3.B2 <> 0) OR ("DB_ALARM".OP3.B3 <> 0) OR ("DB_ALARM".OP3.B4 <> 0) OR ("DB_ALARM".OP3.B5 <> 0) OR ("DB_ALARM".OP3.B6 <> 0) OR ("DB_ALARM".OP3.B7 <> 0) OR ("DB_ALARM".OP3.B8 <> 0) OR ("DB_ALARM".OP3.M_8 <> 0) OR ("DB_ALARM".OP3.M_9 <> 0) OR ("DB_ALARM".OP3.M_10 <> 0) OR ("DB_ALARM".OP3.M_11 <> 0) OR ("DB_ALARM".OP3.M_12 <> 0) OR ("DB_ALARM".OP3.M_13 <> 0) OR ("DB_ALARM".OP3.M_14 <> 0) OR ("DB_ALARM".OP3.M_15 <> 0) OR (%DB100.DBB64 <> 0) OR (%DB100.DBB65 <> 0);
   #OP_3_E := #fc_op_3_alrm;
END_REGION

REGION Network 6: OP_1_WRONG
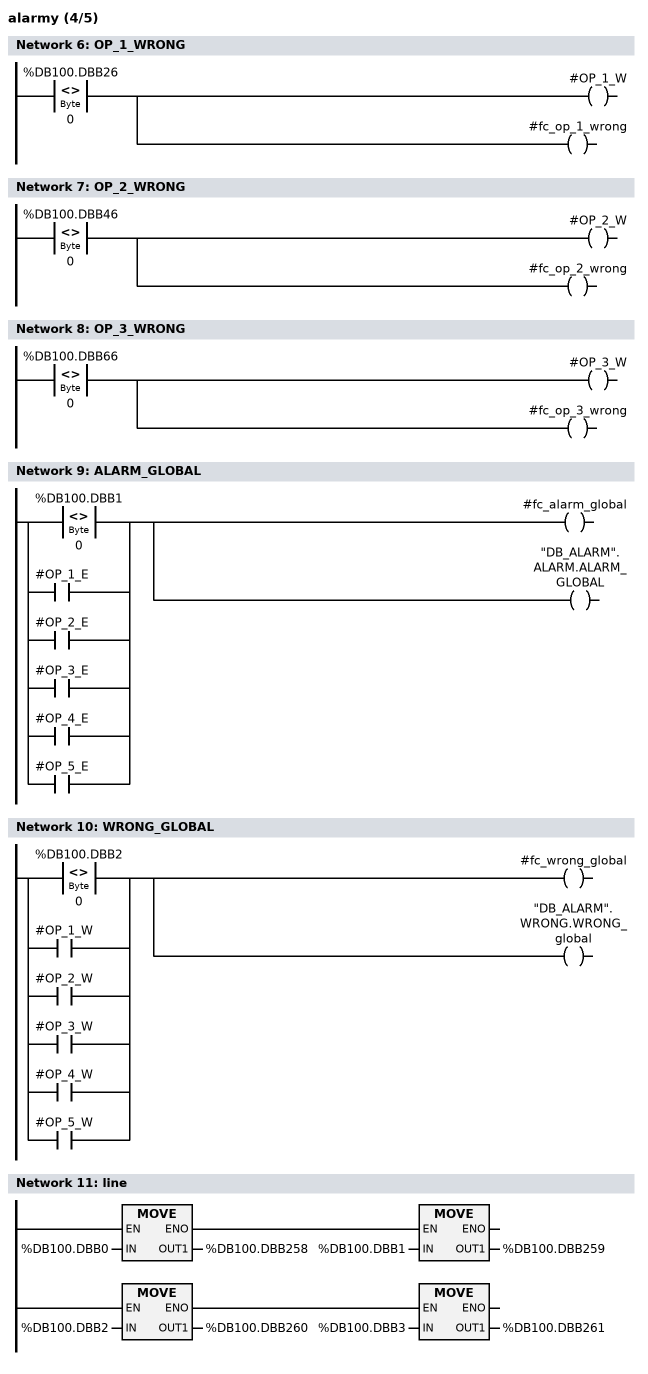
   RUNG wire#powerrail
      { S7_Templates := "SrcType := Byte" } NE_Contact(in1 := %DB100.DBB26, in2 := 0)
      wire#w1
      Coil( #OP_1_W )
   END_RUNG
   RUNG wire#w1
      Coil( #fc_op_1_wrong )
   END_RUNG
   // the same network as SCL:
   #OP_1_W := %DB100.DBB26 <> 0;
   #fc_op_1_wrong := #OP_1_W;
END_REGION

REGION Network 7: OP_2_WRONG
   RUNG wire#powerrail
      { S7_Templates := "SrcType := Byte" } NE_Contact(in1 := %DB100.DBB46, in2 := 0)
      wire#w1
      Coil( #OP_2_W )
   END_RUNG
   RUNG wire#w1
      Coil( #fc_op_2_wrong )
   END_RUNG
   // the same network as SCL:
   #OP_2_W := %DB100.DBB46 <> 0;
   #fc_op_2_wrong := #OP_2_W;
END_REGION

REGION Network 8: OP_3_WRONG
   RUNG wire#powerrail
      { S7_Templates := "SrcType := Byte" } NE_Contact(in1 := %DB100.DBB66, in2 := 0)
      wire#w1
      Coil( #OP_3_W )
   END_RUNG
   RUNG wire#w1
      Coil( #fc_op_3_wrong )
   END_RUNG
   // the same network as SCL:
   #OP_3_W := %DB100.DBB66 <> 0;
   #fc_op_3_wrong := #OP_3_W;
END_REGION

REGION Network 9: ALARM_GLOBAL
   RUNG wire#powerrail
      { S7_Templates := "SrcType := Byte" } NE_Contact(in1 := %DB100.DBB1, in2 := 0)
      wire#w1
      Coil( #fc_alarm_global )
   END_RUNG
   RUNG wire#powerrail
      Contact( #OP_1_E )
   END_RUNG wire#w1
   RUNG wire#powerrail
      Contact( #OP_2_E )
   END_RUNG wire#w1
   RUNG wire#powerrail
      Contact( #OP_3_E )
   END_RUNG wire#w1
   RUNG wire#powerrail
      Contact( #OP_4_E )
   END_RUNG wire#w1
   RUNG wire#powerrail
      Contact( #OP_5_E )
   END_RUNG wire#w1
   RUNG wire#w1
      Coil( "DB_ALARM".ALARM.ALARM_GLOBAL )
   END_RUNG
   // the same network as SCL:
   #fc_alarm_global := (%DB100.DBB1 <> 0) OR #OP_1_E OR #OP_2_E OR #OP_3_E OR #OP_4_E OR #OP_5_E;
   "DB_ALARM".ALARM.ALARM_GLOBAL := #fc_alarm_global;
END_REGION

REGION Network 10: WRONG_GLOBAL
   RUNG wire#powerrail
      { S7_Templates := "SrcType := Byte" } NE_Contact(in1 := %DB100.DBB2, in2 := 0)
      wire#w1
      Coil( #fc_wrong_global )
   END_RUNG
   RUNG wire#powerrail
      Contact( #OP_1_W )
   END_RUNG wire#w1
   RUNG wire#powerrail
      Contact( #OP_2_W )
   END_RUNG wire#w1
   RUNG wire#powerrail
      Contact( #OP_3_W )
   END_RUNG wire#w1
   RUNG wire#powerrail
      Contact( #OP_4_W )
   END_RUNG wire#w1
   RUNG wire#powerrail
      Contact( #OP_5_W )
   END_RUNG wire#w1
   RUNG wire#w1
      Coil( "DB_ALARM".WRONG.WRONG_global )
   END_RUNG
   // the same network as SCL:
   #fc_wrong_global := (%DB100.DBB2 <> 0) OR #OP_1_W OR #OP_2_W OR #OP_3_W OR #OP_4_W OR #OP_5_W;
   "DB_ALARM".WRONG.WRONG_global := #fc_wrong_global;
END_REGION

REGION Network 11: line
   RUNG wire#powerrail
      Move(in := %DB100.DBB0, out1 => %DB100.DBB258)
      Move(in := %DB100.DBB1, out1 => %DB100.DBB259)
   END_RUNG
   RUNG wire#powerrail
      Move(in := %DB100.DBB2, out1 => %DB100.DBB260)
      Move(in := %DB100.DBB3, out1 => %DB100.DBB261)
   END_RUNG
   // the same network as SCL:
   %DB100.DBB258 := %DB100.DBB0;
   %DB100.DBB259 := %DB100.DBB1;
   %DB100.DBB260 := %DB100.DBB2;
   %DB100.DBB261 := %DB100.DBB3;
END_REGION

REGION Network 12: op_1
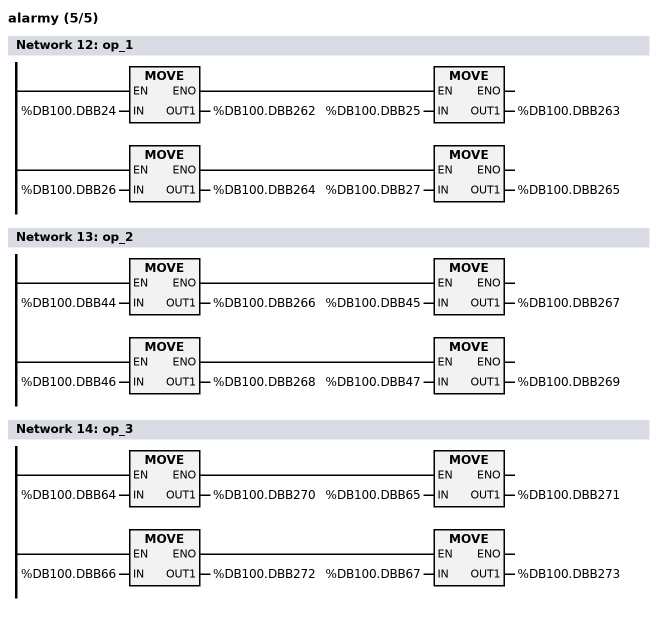
   RUNG wire#powerrail
      Move(in := %DB100.DBB24, out1 => %DB100.DBB262)
      Move(in := %DB100.DBB25, out1 => %DB100.DBB263)
   END_RUNG
   RUNG wire#powerrail
      Move(in := %DB100.DBB26, out1 => %DB100.DBB264)
      Move(in := %DB100.DBB27, out1 => %DB100.DBB265)
   END_RUNG
   // the same network as SCL:
   %DB100.DBB262 := %DB100.DBB24;
   %DB100.DBB263 := %DB100.DBB25;
   %DB100.DBB264 := %DB100.DBB26;
   %DB100.DBB265 := %DB100.DBB27;
END_REGION

REGION Network 13: op_2
   RUNG wire#powerrail
      Move(in := %DB100.DBB44, out1 => %DB100.DBB266)
      Move(in := %DB100.DBB45, out1 => %DB100.DBB267)
   END_RUNG
   RUNG wire#powerrail
      Move(in := %DB100.DBB46, out1 => %DB100.DBB268)
      Move(in := %DB100.DBB47, out1 => %DB100.DBB269)
   END_RUNG
   // the same network as SCL:
   %DB100.DBB266 := %DB100.DBB44;
   %DB100.DBB267 := %DB100.DBB45;
   %DB100.DBB268 := %DB100.DBB46;
   %DB100.DBB269 := %DB100.DBB47;
END_REGION

REGION Network 14: op_3
   RUNG wire#powerrail
      Move(in := %DB100.DBB64, out1 => %DB100.DBB270)
      Move(in := %DB100.DBB65, out1 => %DB100.DBB271)
   END_RUNG
   RUNG wire#powerrail
      Move(in := %DB100.DBB66, out1 => %DB100.DBB272)
      Move(in := %DB100.DBB67, out1 => %DB100.DBB273)
   END_RUNG
   // the same network as SCL:
   %DB100.DBB270 := %DB100.DBB64;
   %DB100.DBB271 := %DB100.DBB65;
   %DB100.DBB272 := %DB100.DBB66;
   %DB100.DBB273 := %DB100.DBB67;
END_REGION

REGION Network 15 (SCL)
   IF "CONTROL_LINE_DB".trig.reset_error_all = TRUE THEN
       // alarm global
       %DB100.DBB0 := 0;
       %DB100.DBB1 := 0;
       // wrong global
       %DB100.DBB2 := 0;
       %DB100.DBB3 := 0;
       // op_0
       // alarm
       %DB100.DBB4 := 0;
       %DB100.DBB5 := 0;
       // wrong
       %DB100.DBB6 := 0;
       %DB100.DBB7 := 0;
       // op_1
       // alarm
       %DB100.DBB24 := 0;
       %DB100.DBB25 := 0;
       // wrong
       %DB100.DBB26 := 0;
       %DB100.DBB27 := 0;
       // op_2
       // alarm
       %DB100.DBB44 := 0;
       %DB100.DBB45 := 0;
       // wrong
       %DB100.DBB46 := 0;
       %DB100.DBB47 := 0;
       // op_3
       // alarm
       %DB100.DBB64 := 0;
       %DB100.DBB65 := 0;
       // wrong
       %DB100.DBB66 := 0;
       %DB100.DBB67 := 0;
       // op_4
       // alarm
       %DB100.DBB84 := 0;
       %DB100.DBB85 := 0;
       // wrong
       %DB100.DBB86 := 0;
       %DB100.DBB87 := 0;
       // op_5
       // alarm
       %DB100.DBB104 := 0;
       %DB100.DBB105 := 0;
       // wrong
       %DB100.DBB106 := 0;
       %DB100.DBB107 := 0;
   END_IF;
END_REGION

REGION Network 16 (SCL)
   //"DB_ALARM".op_0_m_0 := "DB_ALARM".OP0.M_0;
   //"DB_ALARM".op_1_m_0 := "DB_ALARM".OP1.M_0;
   //"DB_ALARM".op_2_m_0 := "DB_ALARM".OP2.A1;
   //"DB_ALARM".op_2_m_1 := "DB_ALARM".OP2.A2;
   //"DB_ALARM".op_2_m_2 := "DB_ALARM".OP2.A3;
   //"DB_ALARM".op_2_m_3 := "DB_ALARM".OP2.A4;
   //"DB_ALARM".op_3_m_0 := "DB_ALARM".OP3.B1;
END_REGION
END_FUNCTION

// folder: STANDARD/CORE/FB_ABMARK_PROFINET

FUNCTION_BLOCK "OVLADANI_LASER"   // FB400, LAD
{ S7_Optimized_Access := 'TRUE' }
VERSION : 0.1
   VAR
      SQCR : Int;
      SQCR_WHILE : Int;
      SET_WHILE : Bool;
      NAZEV_PROGRAMU : String[20];
      DELKA_STRINGU : Int;
      CHAR_K_ZAPISU : Array[0..71] of Char;
   END_VAR
   VAR CONSTANT
      STEP_0 : Int := 0;
      STEP_5 : Int := 5;
      STEP_10 : Int := 10;
      STEP_15 : Int := 15;
      STEP_20 : Int := 20;
      STEP_25 : Int := 25;
      STEP_30 : Int := 30;
      STEP_35 : Int := 35;
      STEP_40 : Int := 40;
      STEP_45 : Int := 45;
      STEP_50 : Int := 50;
      STEP_55 : Int := 55;
      STEP_60 : Int := 60;
      STEP_65 : Int := 65;
      STEP_70 : Int := 70;
      STEP_75 : Int := 75;
      STEP_80 : Int := 80;
      STEP_85 : Int := 85;
      STEP_90 : Int := 90;
      STEP_95 : Int := 95;
      STEP_100 : Int := 100;
   END_VAR
BEGIN

REGION Network 1
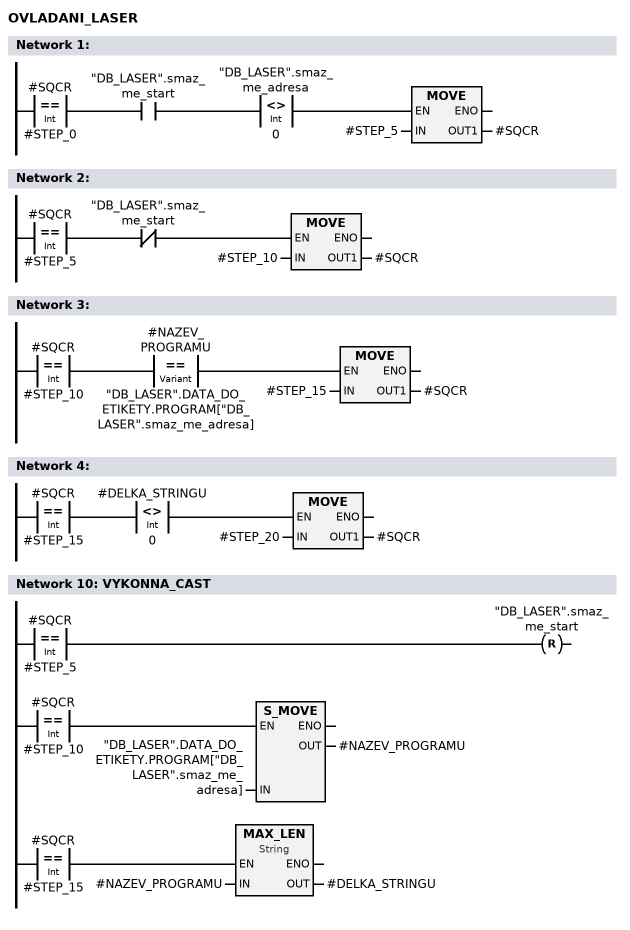
   RUNG wire#powerrail
      { S7_Templates := "SrcType := Int" } EQ_Contact(in1 := #SQCR, in2 := #STEP_0)
      Contact( "DB_LASER".smaz_me_start )
      { S7_Templates := "SrcType := Int" } NE_Contact(in1 := "DB_LASER".smaz_me_adresa, in2 := 0)
      Move(in := #STEP_5, out1 => #SQCR)
   END_RUNG
   // the same network as SCL:
   IF (#SQCR = #STEP_0) AND "DB_LASER".smaz_me_start AND ("DB_LASER".smaz_me_adresa <> 0) THEN
       #SQCR := #STEP_5;
   END_IF;
END_REGION

REGION Network 2
   RUNG wire#powerrail
      { S7_Templates := "SrcType := Int" } EQ_Contact(in1 := #SQCR, in2 := #STEP_5)
      I_Contact( "DB_LASER".smaz_me_start )
      Move(in := #STEP_10, out1 => #SQCR)
   END_RUNG
   // the same network as SCL:
   IF (#SQCR = #STEP_5) AND NOT "DB_LASER".smaz_me_start THEN #SQCR := #STEP_10; END_IF;
END_REGION

REGION Network 3
   RUNG wire#powerrail
      { S7_Templates := "SrcType := Int" } EQ_Contact(in1 := #SQCR, in2 := #STEP_10)
      { S7_Templates := "SrcType := Variant" } EQ_Contact(in1 := #NAZEV_PROGRAMU, in2 := "DB_LASER".DATA_DO_ETIKETY.PROGRAM["DB_LASER".smaz_me_adresa])
      Move(in := #STEP_15, out1 => #SQCR)
   END_RUNG
   // the same network as SCL:
   IF (#SQCR = #STEP_10) AND (#NAZEV_PROGRAMU = "DB_LASER".DATA_DO_ETIKETY.PROGRAM["DB_LASER".smaz_me_adresa]) THEN
       #SQCR := #STEP_15;
   END_IF;
END_REGION

REGION Network 4
   RUNG wire#powerrail
      { S7_Templates := "SrcType := Int" } EQ_Contact(in1 := #SQCR, in2 := #STEP_15)
      { S7_Templates := "SrcType := Int" } NE_Contact(in1 := #DELKA_STRINGU, in2 := 0)
      Move(in := #STEP_20, out1 => #SQCR)
   END_RUNG
   // the same network as SCL:
   IF (#SQCR = #STEP_15) AND (#DELKA_STRINGU <> 0) THEN #SQCR := #STEP_20; END_IF;
END_REGION

REGION Network 5: STEP_20 SCL NETVORK X
END_REGION

REGION Network 10: VYKONNA_CAST
   IF #SQCR = #STEP_5 THEN "DB_LASER".smaz_me_start := FALSE; END_IF;
   IF #SQCR = #STEP_10 THEN
       #NAZEV_PROGRAMU := "DB_LASER".DATA_DO_ETIKETY.PROGRAM["DB_LASER".smaz_me_adresa];
   END_IF;
   IF #SQCR = #STEP_15 THEN MAX_LEN(in := #NAZEV_PROGRAMU, out => #DELKA_STRINGU); END_IF;
END_REGION

REGION Network 12 (SCL)
   IF #SQCR = #STEP_20 THEN
       // zapsani počátečního znaku 
       #CHAR_K_ZAPISU[0] := "DB_LASER".DATA_DO_DAT.ZAVORKA_P;



       // vytvoření prdelky k názvu programu z laseru
       #CHAR_K_ZAPISU[#DELKA_STRINGU + 1] := "DB_LASER".DATA_DO_DAT.XLP[0];
       #CHAR_K_ZAPISU[#DELKA_STRINGU + 2] := "DB_LASER".DATA_DO_DAT.XLP[1];
       #CHAR_K_ZAPISU[#DELKA_STRINGU + 3] := "DB_LASER".DATA_DO_DAT.XLP[2];
       #CHAR_K_ZAPISU[#DELKA_STRINGU + 4] := "DB_LASER".DATA_DO_DAT.XLP[3];
       #CHAR_K_ZAPISU[#DELKA_STRINGU + 5] := "DB_LASER".DATA_DO_DAT.ZAVORKA_P;

       // dinamický zápis názvu podle délky stringu 
       WHILE #SET_WHILE DO
           IF #SQCR_WHILE > #DELKA_STRINGU THEN
               #SQCR_WHILE := 0;
               #SET_WHILE := FALSE;
               #SQCR := #STEP_25;
           ELSE
               #SQCR_WHILE := #SQCR_WHILE + 1;
           END_IF;
           #CHAR_K_ZAPISU[#SQCR_WHILE + 1] := #NAZEV_PROGRAMU[#SQCR_WHILE];
       END_WHILE;

   END_IF;
END_REGION
END_FUNCTION_BLOCK

FUNCTION "DATA_R/W" : Void   // FC400, SCL
{ S7_Optimized_Access := 'TRUE' }
VERSION : 0.1
BEGIN
   IF "DB_DATA_LASER".READ = TRUE THEN
       "DB_DATA_LASER".LASER_DATA_READ[0] := "RESPONSE_DATA_FIELD_0";
       "DB_DATA_LASER".LASER_DATA_READ[1] := "RESPONSE_DATA_FIELD_1";
       "DB_DATA_LASER".LASER_DATA_READ[2] := "RESPONSE_DATA_FIELD_2";
       "DB_DATA_LASER".LASER_DATA_READ[3] := "RESPONSE_DATA_FIELD_3";
       "DB_DATA_LASER".LASER_DATA_READ[4] := "RESPONSE_DATA_FIELD_4";
       "DB_DATA_LASER".LASER_DATA_READ[5] := "RESPONSE_DATA_FIELD_5";
       "DB_DATA_LASER".LASER_DATA_READ[6] := "RESPONSE_DATA_FIELD_6";
       "DB_DATA_LASER".LASER_DATA_READ[7] := "RESPONSE_DATA_FIELD_7";
       "DB_DATA_LASER".LASER_DATA_READ[8] := "RESPONSE_DATA_FIELD_8";
       "DB_DATA_LASER".LASER_DATA_READ[9] := "RESPONSE_DATA_FIELD_9";
       "DB_DATA_LASER".LASER_DATA_READ[10] := "RESPONSE_DATA_FIELD_10";
       "DB_DATA_LASER".LASER_DATA_READ[11] := "RESPONSE_DATA_FIELD_11";
       "DB_DATA_LASER".LASER_DATA_READ[12] := "RESPONSE_DATA_FIELD_12";
       "DB_DATA_LASER".LASER_DATA_READ[13] := "RESPONSE_DATA_FIELD_13";
       "DB_DATA_LASER".LASER_DATA_READ[14] := "RESPONSE_DATA_FIELD_14";
       "DB_DATA_LASER".LASER_DATA_READ[15] := "RESPONSE_DATA_FIELD_15";
       "DB_DATA_LASER".LASER_DATA_READ[16] := "RESPONSE_DATA_FIELD_16";
       "DB_DATA_LASER".LASER_DATA_READ[17] := "RESPONSE_DATA_FIELD_17";
       "DB_DATA_LASER".LASER_DATA_READ[18] := "RESPONSE_DATA_FIELD_18";
       "DB_DATA_LASER".LASER_DATA_READ[19] := "RESPONSE_DATA_FIELD_19";
       "DB_DATA_LASER".LASER_DATA_READ[20] := "RESPONSE_DATA_FIELD_20";
       "DB_DATA_LASER".LASER_DATA_READ[21] := "RESPONSE_DATA_FIELD_21";
       "DB_DATA_LASER".LASER_DATA_READ[22] := "RESPONSE_DATA_FIELD_22";
       "DB_DATA_LASER".LASER_DATA_READ[23] := "RESPONSE_DATA_FIELD_23";
       "DB_DATA_LASER".LASER_DATA_READ[24] := "RESPONSE_DATA_FIELD_24";
       "DB_DATA_LASER".LASER_DATA_READ[25] := "RESPONSE_DATA_FIELD_25";
       "DB_DATA_LASER".LASER_DATA_READ[26] := "RESPONSE_DATA_FIELD_26";
       "DB_DATA_LASER".LASER_DATA_READ[27] := "RESPONSE_DATA_FIELD_27";
       "DB_DATA_LASER".LASER_DATA_READ[28] := "RESPONSE_DATA_FIELD_28";
       "DB_DATA_LASER".LASER_DATA_READ[29] := "RESPONSE_DATA_FIELD_29";
       "DB_DATA_LASER".LASER_DATA_READ[30] := "RESPONSE_DATA_FIELD_30";
       "DB_DATA_LASER".LASER_DATA_READ[31] := "RESPONSE_DATA_FIELD_31";
       "DB_DATA_LASER".LASER_DATA_READ[32] := "RESPONSE_DATA_FIELD_32";
       "DB_DATA_LASER".LASER_DATA_READ[33] := "RESPONSE_DATA_FIELD_33";
       "DB_DATA_LASER".LASER_DATA_READ[34] := "RESPONSE_DATA_FIELD_34";
       "DB_DATA_LASER".LASER_DATA_READ[35] := "RESPONSE_DATA_FIELD_35";
       "DB_DATA_LASER".LASER_DATA_READ[36] := "RESPONSE_DATA_FIELD_36";
       "DB_DATA_LASER".LASER_DATA_READ[37] := "RESPONSE_DATA_FIELD_37";
       "DB_DATA_LASER".LASER_DATA_READ[38] := "RESPONSE_DATA_FIELD_38";
       "DB_DATA_LASER".LASER_DATA_READ[39] := "RESPONSE_DATA_FIELD_39";
       "DB_DATA_LASER".LASER_DATA_READ[40] := "RESPONSE_DATA_FIELD_40";
       "DB_DATA_LASER".LASER_DATA_READ[41] := "RESPONSE_DATA_FIELD_41";
       "DB_DATA_LASER".LASER_DATA_READ[42] := "RESPONSE_DATA_FIELD_42";
       "DB_DATA_LASER".LASER_DATA_READ[43] := "RESPONSE_DATA_FIELD_43";
       "DB_DATA_LASER".LASER_DATA_READ[44] := "RESPONSE_DATA_FIELD_44";
       "DB_DATA_LASER".LASER_DATA_READ[45] := "RESPONSE_DATA_FIELD_45";
       "DB_DATA_LASER".LASER_DATA_READ[46] := "RESPONSE_DATA_FIELD_46";
       "DB_DATA_LASER".LASER_DATA_READ[47] := "RESPONSE_DATA_FIELD_47";
       "DB_DATA_LASER".LASER_DATA_READ[48] := "RESPONSE_DATA_FIELD_48";
       "DB_DATA_LASER".LASER_DATA_READ[49] := "RESPONSE_DATA_FIELD_49";
       "DB_DATA_LASER".LASER_DATA_READ[50] := "RESPONSE_DATA_FIELD_50";
       "DB_DATA_LASER".LASER_DATA_READ[51] := "RESPONSE_DATA_FIELD_51";
       "DB_DATA_LASER".LASER_DATA_READ[52] := "RESPONSE_DATA_FIELD_52";
       "DB_DATA_LASER".LASER_DATA_READ[53] := "RESPONSE_DATA_FIELD_53";
       "DB_DATA_LASER".LASER_DATA_READ[54] := "RESPONSE_DATA_FIELD_54";
       "DB_DATA_LASER".LASER_DATA_READ[55] := "RESPONSE_DATA_FIELD_55";
       "DB_DATA_LASER".LASER_DATA_READ[56] := "RESPONSE_DATA_FIELD_56";
       "DB_DATA_LASER".LASER_DATA_READ[57] := "RESPONSE_DATA_FIELD_57";
       "DB_DATA_LASER".LASER_DATA_READ[58] := "RESPONSE_DATA_FIELD_58";
       "DB_DATA_LASER".LASER_DATA_READ[59] := "RESPONSE_DATA_FIELD_59";
       "DB_DATA_LASER".LASER_DATA_READ[60] := "RESPONSE_DATA_FIELD_60";
       "DB_DATA_LASER".LASER_DATA_READ[61] := "RESPONSE_DATA_FIELD_61";
       "DB_DATA_LASER".LASER_DATA_READ[62] := "RESPONSE_DATA_FIELD_62";
       "DB_DATA_LASER".LASER_DATA_READ[63] := "RESPONSE_DATA_FIELD_63";
       "DB_DATA_LASER".LASER_DATA_READ[64] := "RESPONSE_DATA_FIELD_64";
       "DB_DATA_LASER".LASER_DATA_READ[65] := "RESPONSE_DATA_FIELD_65";
       "DB_DATA_LASER".LASER_DATA_READ[66] := "RESPONSE_DATA_FIELD_66";
       "DB_DATA_LASER".LASER_DATA_READ[67] := "RESPONSE_DATA_FIELD_67";
       "DB_DATA_LASER".LASER_DATA_READ[68] := "RESPONSE_DATA_FIELD_68";
       "DB_DATA_LASER".LASER_DATA_READ[69] := "RESPONSE_DATA_FIELD_69";
       "DB_DATA_LASER".LASER_DATA_READ[70] := "RESPONSE_DATA_FIELD_70";
       "DB_DATA_LASER".LASER_DATA_READ[71] := "RESPONSE_DATA_FIELD_71";

       "DB_DATA_LASER".READ := FALSE;
   END_IF;
    (*   
   IF "DB_DATA_LASER".WRITE = TRUE THEN
       "REQUEST_DATA_FIELC_BYTE_0" := "DB_DATA_LASER".LASER_DATA_WRITE[0];
       "REQUEST_DATA_FIELC_BYTE_1" := "DB_DATA_LASER".LASER_DATA_WRITE[1];
       "REQUEST_DATA_FIELC_BYTE_2" := "DB_DATA_LASER".LASER_DATA_WRITE[2];
       "REQUEST_DATA_FIELC_BYTE_3" := "DB_DATA_LASER".LASER_DATA_WRITE[3];
       "REQUEST_DATA_FIELC_BYTE_4" := "DB_DATA_LASER".LASER_DATA_WRITE[4];
       "REQUEST_DATA_FIELC_BYTE_5" := "DB_DATA_LASER".LASER_DATA_WRITE[5];
       "REQUEST_DATA_FIELC_BYTE_6" := "DB_DATA_LASER".LASER_DATA_WRITE[6];
       "REQUEST_DATA_FIELC_BYTE_7" := "DB_DATA_LASER".LASER_DATA_WRITE[7];
       "REQUEST_DATA_FIELC_BYTE_8" := "DB_DATA_LASER".LASER_DATA_WRITE[8];
       "REQUEST_DATA_FIELC_BYTE_9" := "DB_DATA_LASER".LASER_DATA_WRITE[9];
       "REQUEST_DATA_FIELC_BYTE_10" := "DB_DATA_LASER".LASER_DATA_WRITE[10];
       "REQUEST_DATA_FIELC_BYTE_11" := "DB_DATA_LASER".LASER_DATA_WRITE[11];
       "REQUEST_DATA_FIELC_BYTE_12" := "DB_DATA_LASER".LASER_DATA_WRITE[12];
       "REQUEST_DATA_FIELC_BYTE_13" := "DB_DATA_LASER".LASER_DATA_WRITE[13];
       "REQUEST_DATA_FIELC_BYTE_14" := "DB_DATA_LASER".LASER_DATA_WRITE[14];
       "REQUEST_DATA_FIELC_BYTE_15" := "DB_DATA_LASER".LASER_DATA_WRITE[15];
       "REQUEST_DATA_FIELC_BYTE_16" := "DB_DATA_LASER".LASER_DATA_WRITE[16];
       "REQUEST_DATA_FIELC_BYTE_17" := "DB_DATA_LASER".LASER_DATA_WRITE[17];
       "REQUEST_DATA_FIELC_BYTE_18" := "DB_DATA_LASER".LASER_DATA_WRITE[18];
       "REQUEST_DATA_FIELC_BYTE_19" := "DB_DATA_LASER".LASER_DATA_WRITE[19];
       "REQUEST_DATA_FIELC_BYTE_20" := "DB_DATA_LASER".LASER_DATA_WRITE[20];
       "REQUEST_DATA_FIELC_BYTE_21" := "DB_DATA_LASER".LASER_DATA_WRITE[21];
       "REQUEST_DATA_FIELC_BYTE_22" := "DB_DATA_LASER".LASER_DATA_WRITE[22];
       "REQUEST_DATA_FIELC_BYTE_23" := "DB_DATA_LASER".LASER_DATA_WRITE[23];
       "REQUEST_DATA_FIELC_BYTE_24" := "DB_DATA_LASER".LASER_DATA_WRITE[24];
       "REQUEST_DATA_FIELC_BYTE_25" := "DB_DATA_LASER".LASER_DATA_WRITE[25];
       "REQUEST_DATA_FIELC_BYTE_26" := "DB_DATA_LASER".LASER_DATA_WRITE[26];
       "REQUEST_DATA_FIELC_BYTE_27" := "DB_DATA_LASER".LASER_DATA_WRITE[27];
       "REQUEST_DATA_FIELC_BYTE_28" := "DB_DATA_LASER".LASER_DATA_WRITE[28];
       "REQUEST_DATA_FIELC_BYTE_29" := "DB_DATA_LASER".LASER_DATA_WRITE[29];
       "REQUEST_DATA_FIELC_BYTE_30" := "DB_DATA_LASER".LASER_DATA_WRITE[30];
       "REQUEST_DATA_FIELC_BYTE_31" := "DB_DATA_LASER".LASER_DATA_WRITE[31];
       "REQUEST_DATA_FIELC_BYTE_32" := "DB_DATA_LASER".LASER_DATA_WRITE[32];
       "REQUEST_DATA_FIELC_BYTE_33" := "DB_DATA_LASER".LASER_DATA_WRITE[33];
       "REQUEST_DATA_FIELC_BYTE_34" := "DB_DATA_LASER".LASER_DATA_WRITE[34];
       "REQUEST_DATA_FIELC_BYTE_35" := "DB_DATA_LASER".LASER_DATA_WRITE[35];
       "REQUEST_DATA_FIELC_BYTE_36" := "DB_DATA_LASER".LASER_DATA_WRITE[36];
       "REQUEST_DATA_FIELC_BYTE_37" := "DB_DATA_LASER".LASER_DATA_WRITE[37];
       "REQUEST_DATA_FIELC_BYTE_38" := "DB_DATA_LASER".LASER_DATA_WRITE[38];
       "REQUEST_DATA_FIELC_BYTE_39" := "DB_DATA_LASER".LASER_DATA_WRITE[39];
       "REQUEST_DATA_FIELC_BYTE_40" := "DB_DATA_LASER".LASER_DATA_WRITE[40];
       "REQUEST_DATA_FIELC_BYTE_41" := "DB_DATA_LASER".LASER_DATA_WRITE[41];
       "REQUEST_DATA_FIELC_BYTE_42" := "DB_DATA_LASER".LASER_DATA_WRITE[42];
       "REQUEST_DATA_FIELC_BYTE_43" := "DB_DATA_LASER".LASER_DATA_WRITE[43];
       "REQUEST_DATA_FIELC_BYTE_44" := "DB_DATA_LASER".LASER_DATA_WRITE[44];
       "REQUEST_DATA_FIELC_BYTE_45" := "DB_DATA_LASER".LASER_DATA_WRITE[45];
       "REQUEST_DATA_FIELC_BYTE_46" := "DB_DATA_LASER".LASER_DATA_WRITE[46];
       "REQUEST_DATA_FIELC_BYTE_47" := "DB_DATA_LASER".LASER_DATA_WRITE[47];
       "REQUEST_DATA_FIELC_BYTE_48" := "DB_DATA_LASER".LASER_DATA_WRITE[48];
       "REQUEST_DATA_FIELC_BYTE_49" := "DB_DATA_LASER".LASER_DATA_WRITE[49];
       "REQUEST_DATA_FIELC_BYTE_50" := "DB_DATA_LASER".LASER_DATA_WRITE[50];
       "REQUEST_DATA_FIELC_BYTE_51" := "DB_DATA_LASER".LASER_DATA_WRITE[51];
       "REQUEST_DATA_FIELC_BYTE_52" := "DB_DATA_LASER".LASER_DATA_WRITE[52];
       "REQUEST_DATA_FIELC_BYTE_53" := "DB_DATA_LASER".LASER_DATA_WRITE[53];
       "REQUEST_DATA_FIELC_BYTE_54" := "DB_DATA_LASER".LASER_DATA_WRITE[54];
       "REQUEST_DATA_FIELC_BYTE_55" := "DB_DATA_LASER".LASER_DATA_WRITE[55];
       "REQUEST_DATA_FIELC_BYTE_56" := "DB_DATA_LASER".LASER_DATA_WRITE[56];
       "REQUEST_DATA_FIELC_BYTE_57" := "DB_DATA_LASER".LASER_DATA_WRITE[57];
       "REQUEST_DATA_FIELC_BYTE_58" := "DB_DATA_LASER".LASER_DATA_WRITE[58];
       "REQUEST_DATA_FIELC_BYTE_59" := "DB_DATA_LASER".LASER_DATA_WRITE[59];
       "REQUEST_DATA_FIELC_BYTE_60" := "DB_DATA_LASER".LASER_DATA_WRITE[60];
       "REQUEST_DATA_FIELC_BYTE_61" := "DB_DATA_LASER".LASER_DATA_WRITE[61];
       "REQUEST_DATA_FIELC_BYTE_62" := "DB_DATA_LASER".LASER_DATA_WRITE[62];
       "REQUEST_DATA_FIELC_BYTE_63" := "DB_DATA_LASER".LASER_DATA_WRITE[63];
       "REQUEST_DATA_FIELC_BYTE_64" := "DB_DATA_LASER".LASER_DATA_WRITE[64];
       "REQUEST_DATA_FIELC_BYTE_65" := "DB_DATA_LASER".LASER_DATA_WRITE[65];
       "REQUEST_DATA_FIELC_BYTE_66" := "DB_DATA_LASER".LASER_DATA_WRITE[66];
       "REQUEST_DATA_FIELC_BYTE_67" := "DB_DATA_LASER".LASER_DATA_WRITE[67];
       "REQUEST_DATA_FIELC_BYTE_68" := "DB_DATA_LASER".LASER_DATA_WRITE[68];
       "REQUEST_DATA_FIELC_BYTE_69" := "DB_DATA_LASER".LASER_DATA_WRITE[69];
       "REQUEST_DATA_FIELC_BYTE_70" := "DB_DATA_LASER".LASER_DATA_WRITE[70];
       "REQUEST_DATA_FIELC_BYTE_71" := "DB_DATA_LASER".LASER_DATA_WRITE[71];

       "DB_DATA_LASER".WRITE := FALSE;
   END_IF;
   *)
END_FUNCTION

// folder: STANDARD/LINE

FUNCTION_BLOCK "CONTROL_LINE"   // FB7, LAD
{ S7_Optimized_Access := 'TRUE' }
VERSION : 0.1
   VAR
      TIMER_reset : TON_TIME;
      P_TRIG_INICIAL : Bool;
      P_TRIG_RESET : Bool;
      AUTOMAT : "SENSOR";
      MANUAL : "SENSOR";
      SENSOR_3 : "SENSOR";
      SENSOR_4 : "SENSOR";
      SENSOR_5 : "SENSOR";
      SENSOR_6 : "SENSOR";
      SENSOR_7 : "SENSOR";
      SENSOR_8 : "SENSOR";
      SENSOR_9 : "SENSOR";
      SENSOR_10 : "SENSOR";
      SENSOR_11 : "SENSOR";
      dvere_L_A : "SENSOR";
      dvere_L_B : "SENSOR";
      dvere_P_A : "SENSOR";
      dvere_P_B : "SENSOR";
      SEN_STRUCT : Struct
         AUTOMAT : Bool;
         AUTOMAT_NEG : Bool;
         MANUAL : Bool;
         MANUAL_NEG : Bool;
         SENSOR_TLAKU : Bool;
         SENSOR_TLAKU_NEG : Bool;
         power : Bool;
         power_neg : Bool;
         safety : Bool;
         safety_neg : Bool;
         s_10 : Bool;
         TLA_STOP : Bool;
         TLA_STOP_NEG : Bool;
         TLA_START : Bool;
         TLA_START_NEG : Bool;
         TLA_KVIT : Bool;
         TLA_KVIT_NEG : Bool;
         s_17 : Bool;
         S19 : Bool;
         L1_OK : Bool;
         L1_NOT_OK : Bool;
         L2_OK : Bool;
         L2_NOT_OK : Bool;
         L3_OK : Bool;
         L3_NOT_OK : Bool;
         dvere_L_A : Bool;
         dvere_L_B : Bool;
         dvere_P_A : Bool;
         dvere_P_B : Bool;
         S30 : Bool;
         S31 : Bool;
         LASER_MEMOR : Bool;
      END_STRUCT;
      "M" : Struct
         P_TRIK_hmi_manual : Bool;
         p_trig_hmi_automat : Bool;
         N_TRIG_REZIM : Bool;
         M_4 : Bool;
         hlaseni_chyby : Bool;
         M_6 : Bool;
         M_7 : Bool;
         M_8 : Bool;
         M_9 : Bool;
         p_Trig_al : Bool;
         n_trig_al : Bool;
         p_trig_wro : Bool;
         n_trig_wro : Bool;
         M_14 : Bool;
         M_15 : Bool;
         N_TRIG_MANUAL : Bool;
         M_17 : Bool;
         M_18 : Bool;
         M_19 : Bool;
         M_20 : Bool;
         M_21 : Bool;
         M_22 : Bool;
         M_23 : Bool;
         M_24 : Bool;
         M_25 : Bool;
         M_26 : Bool;
         M_27 : Bool;
         M_28 : Bool;
         M_29 : Bool;
         M_30 : Bool;
         M_31 : Bool;
         M_32 : Bool;
      END_STRUCT;
      trig : Struct
         reset_error_all : Bool;
         TRIG_FOR_OP_4_AUTOMAT : Bool;
         t_3 : Bool;
         t_4 : Bool;
         t_5 : Bool;
         t_6 : Bool;
         t_7 : Bool;
         t_8 : Bool;
      END_STRUCT;
      SQCR : Int;
      job_mailbox : Array[0..3] of Word;
      n_trig_res_auit : Bool;
      inicial_control : TON_TIME;
      SQCR_SAFETY : Int;
      n_trig_RESET_AUT : Bool;
      P_TRIG_RESET_SAFETY : Bool;
      air : TON_TIME;
      HMI_ALARM : Int;
   END_VAR
   VAR_TEMP
      "string" : String;
      smaz_me : Bool;
      majak_green_s1 : Bool;
      majak_red_s1 : Bool;
      majak_yelou_s1 : Bool;
      majak_blue_s1 : Bool;
      majak_orange_s1 : Bool;
      majak_green_s2 : Bool;
      majak_red_s2 : Bool;
      majak_yelou_s2 : Bool;
      majak_blue_s2 : Bool;
      majak_orange_s2 : Bool;
      majak_green_s3 : Bool;
      majak_red_s3 : Bool;
      majak_yelou_s3 : Bool;
      majak_blue_s3 : Bool;
      majak_orange_s3 : Bool;
      majak_green_s4 : Bool;
      majak_red_s4 : Bool;
      majak_yelou_s4 : Bool;
      majak_blue_s4 : Bool;
      majak_orange_s4 : Bool;
      majak_green_s5 : Bool;
      majak_red_s5 : Bool;
      majak_yelou_s5 : Bool;
      majak_blue_s5 : Bool;
      majak_orange_s5 : Bool;
   END_VAR
   VAR CONSTANT
      STEP_0_FIRST_START : Int := 0;
      STEP_3 : Int := 3;
      STEP_5 : Int := 5;
      STEP_10 : Int := 10;
      STEP_15 : Int := 15;
      STEP_20 : Int := 20;
      STEP_25 : Int := 25;
      STEP_27 : Int := 27;
      STEP_30 : Int := 30;
      STEP_35 : Int := 35;
      STEP_40 : Int := 40;
      STEP_45 : Int := 45;
      STEP_48 : Int := 48;
      STEP_50 : Int := 50;
      STEP_52 : Int := 52;
      STEP_55 : Int := 55;
      STEP_60 : Int := 60;
      STEP_65 : Int := 65;
      STEP_70 : Int := 70;
      STEP_75 : Int := 75;
      STEP_80 : Int := 80;
      STEP_85 : Int := 85;
      STEP_90 : Int := 90;
      STEP_95 : Int := 95;
      STEP_100 : Int := 100;
      STEO_105 : Int := 105;
   END_VAR
   VAR_TEMP   // added for the SCL form of the ladder/FBD networks
      _w1 : Bool;
      _w2 : Bool;
      _w3 : Bool;
      _w4 : Bool;
      _w5 : Bool;
   END_VAR
BEGIN

REGION Network 1 (SCL)
   // SET  BASIC ELEMENTS
   // odpojení nepoužívaných kontaktů
   "LOG_0" := 0;
   "LOG_1" := 1;
   "SMAZ_ME_0" := 0;
   "SMAZ_ME_1" := 1;
END_REGION

REGION Network 2: SENSORS
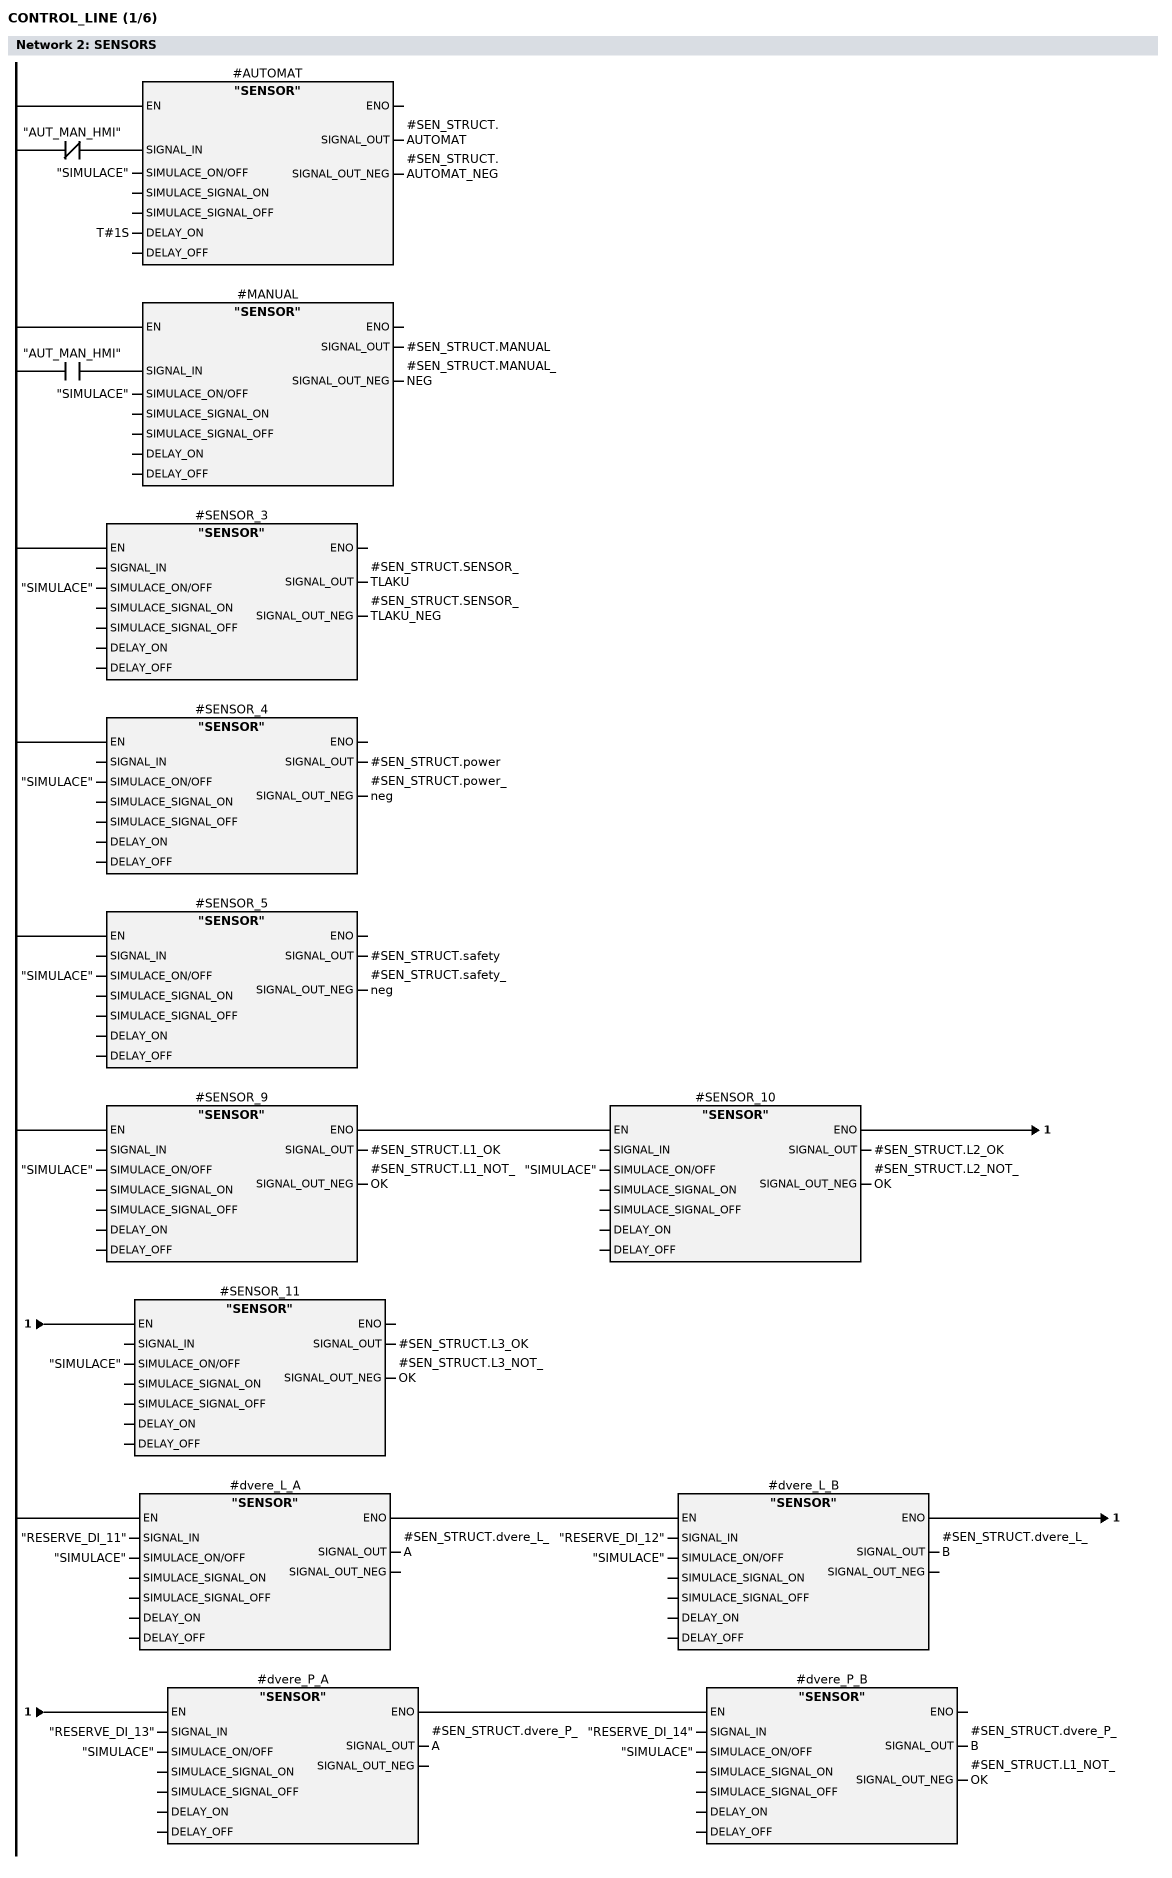
   RUNG wire#powerrail
      #AUTOMAT(SIGNAL_IN := wire#w1, "SIMULACE_ON/OFF" := "SIMULACE", SIMULACE_SIGNAL_ON :=, SIMULACE_SIGNAL_OFF :=, DELAY_ON := T#1S, DELAY_OFF :=, SIGNAL_OUT => #SEN_STRUCT.AUTOMAT, SIGNAL_OUT_NEG => #SEN_STRUCT.AUTOMAT_NEG)
   END_RUNG
   RUNG wire#powerrail
      I_Contact( "AUT_MAN_HMI" )
   END_RUNG wire#w1
   RUNG wire#powerrail
      #MANUAL(SIGNAL_IN := wire#w2, "SIMULACE_ON/OFF" := "SIMULACE", SIMULACE_SIGNAL_ON :=, SIMULACE_SIGNAL_OFF :=, DELAY_ON :=, DELAY_OFF :=, SIGNAL_OUT => #SEN_STRUCT.MANUAL, SIGNAL_OUT_NEG => #SEN_STRUCT.MANUAL_NEG)
   END_RUNG
   RUNG wire#powerrail
      Contact( "AUT_MAN_HMI" )
   END_RUNG wire#w2
   RUNG wire#powerrail
      #SENSOR_3(SIGNAL_IN :=, "SIMULACE_ON/OFF" := "SIMULACE", SIMULACE_SIGNAL_ON :=, SIMULACE_SIGNAL_OFF :=, DELAY_ON :=, DELAY_OFF :=, SIGNAL_OUT => #SEN_STRUCT.SENSOR_TLAKU, SIGNAL_OUT_NEG => #SEN_STRUCT.SENSOR_TLAKU_NEG)
   END_RUNG
   RUNG wire#powerrail
      #SENSOR_4(SIGNAL_IN :=, "SIMULACE_ON/OFF" := "SIMULACE", SIMULACE_SIGNAL_ON :=, SIMULACE_SIGNAL_OFF :=, DELAY_ON :=, DELAY_OFF :=, SIGNAL_OUT => #SEN_STRUCT.power, SIGNAL_OUT_NEG => #SEN_STRUCT.power_neg)
   END_RUNG
   RUNG wire#powerrail
      #SENSOR_5(SIGNAL_IN :=, "SIMULACE_ON/OFF" := "SIMULACE", SIMULACE_SIGNAL_ON :=, SIMULACE_SIGNAL_OFF :=, DELAY_ON :=, DELAY_OFF :=, SIGNAL_OUT => #SEN_STRUCT.safety, SIGNAL_OUT_NEG => #SEN_STRUCT.safety_neg)
   END_RUNG
   RUNG wire#powerrail
      #SENSOR_9(SIGNAL_IN :=, "SIMULACE_ON/OFF" := "SIMULACE", SIMULACE_SIGNAL_ON :=, SIMULACE_SIGNAL_OFF :=, DELAY_ON :=, DELAY_OFF :=, SIGNAL_OUT => #SEN_STRUCT.L1_OK, SIGNAL_OUT_NEG => #SEN_STRUCT.L1_NOT_OK)
      #SENSOR_10(SIGNAL_IN :=, "SIMULACE_ON/OFF" := "SIMULACE", SIMULACE_SIGNAL_ON :=, SIMULACE_SIGNAL_OFF :=, DELAY_ON :=, DELAY_OFF :=, SIGNAL_OUT => #SEN_STRUCT.L2_OK, SIGNAL_OUT_NEG => #SEN_STRUCT.L2_NOT_OK)
      #SENSOR_11(SIGNAL_IN :=, "SIMULACE_ON/OFF" := "SIMULACE", SIMULACE_SIGNAL_ON :=, SIMULACE_SIGNAL_OFF :=, DELAY_ON :=, DELAY_OFF :=, SIGNAL_OUT => #SEN_STRUCT.L3_OK, SIGNAL_OUT_NEG => #SEN_STRUCT.L3_NOT_OK)
   END_RUNG
   RUNG wire#powerrail
      #dvere_L_A(SIGNAL_IN := "RESERVE_DI_11", "SIMULACE_ON/OFF" := "SIMULACE", SIMULACE_SIGNAL_ON :=, SIMULACE_SIGNAL_OFF :=, DELAY_ON :=, DELAY_OFF :=, SIGNAL_OUT => #SEN_STRUCT.dvere_L_A, SIGNAL_OUT_NEG =>)
      #dvere_L_B(SIGNAL_IN := "RESERVE_DI_12", "SIMULACE_ON/OFF" := "SIMULACE", SIMULACE_SIGNAL_ON :=, SIMULACE_SIGNAL_OFF :=, DELAY_ON :=, DELAY_OFF :=, SIGNAL_OUT => #SEN_STRUCT.dvere_L_B, SIGNAL_OUT_NEG =>)
      #dvere_P_A(SIGNAL_IN := "RESERVE_DI_13", "SIMULACE_ON/OFF" := "SIMULACE", SIMULACE_SIGNAL_ON :=, SIMULACE_SIGNAL_OFF :=, DELAY_ON :=, DELAY_OFF :=, SIGNAL_OUT => #SEN_STRUCT.dvere_P_A, SIGNAL_OUT_NEG =>)
      #dvere_P_B(SIGNAL_IN := "RESERVE_DI_14", "SIMULACE_ON/OFF" := "SIMULACE", SIMULACE_SIGNAL_ON :=, SIMULACE_SIGNAL_OFF :=, DELAY_ON :=, DELAY_OFF :=, SIGNAL_OUT => #SEN_STRUCT.dvere_P_B, SIGNAL_OUT_NEG => #SEN_STRUCT.L1_NOT_OK)
   END_RUNG
   // the same network as SCL:
   #AUTOMAT(SIGNAL_IN := NOT "AUT_MAN_HMI",   // "SENSOR"
            "SIMULACE_ON/OFF" := "SIMULACE",
            DELAY_ON := T#1S,
            SIGNAL_OUT => #SEN_STRUCT.AUTOMAT,
            SIGNAL_OUT_NEG => #SEN_STRUCT.AUTOMAT_NEG);
   #MANUAL(SIGNAL_IN := "AUT_MAN_HMI",   // "SENSOR"
           "SIMULACE_ON/OFF" := "SIMULACE",
           SIGNAL_OUT => #SEN_STRUCT.MANUAL,
           SIGNAL_OUT_NEG => #SEN_STRUCT.MANUAL_NEG);
   #SENSOR_3("SIMULACE_ON/OFF" := "SIMULACE",   // "SENSOR"
             SIGNAL_OUT => #SEN_STRUCT.SENSOR_TLAKU,
             SIGNAL_OUT_NEG => #SEN_STRUCT.SENSOR_TLAKU_NEG);
   #SENSOR_4("SIMULACE_ON/OFF" := "SIMULACE",   // "SENSOR"
             SIGNAL_OUT => #SEN_STRUCT.power,
             SIGNAL_OUT_NEG => #SEN_STRUCT.power_neg);
   #SENSOR_5("SIMULACE_ON/OFF" := "SIMULACE",   // "SENSOR"
             SIGNAL_OUT => #SEN_STRUCT.safety,
             SIGNAL_OUT_NEG => #SEN_STRUCT.safety_neg);
   #SENSOR_9("SIMULACE_ON/OFF" := "SIMULACE",   // "SENSOR"
             SIGNAL_OUT => #SEN_STRUCT.L1_OK,
             SIGNAL_OUT_NEG => #SEN_STRUCT.L1_NOT_OK,
             ENO => #_w1);
   #SENSOR_10(EN := #_w1,   // "SENSOR"
              "SIMULACE_ON/OFF" := "SIMULACE",
              SIGNAL_OUT => #SEN_STRUCT.L2_OK,
              SIGNAL_OUT_NEG => #SEN_STRUCT.L2_NOT_OK,
              ENO => #_w2);
   IF #_w2 THEN
       #SENSOR_11("SIMULACE_ON/OFF" := "SIMULACE",   // "SENSOR"
                  SIGNAL_OUT => #SEN_STRUCT.L3_OK,
                  SIGNAL_OUT_NEG => #SEN_STRUCT.L3_NOT_OK);
   END_IF;
   #dvere_L_A(SIGNAL_IN := "RESERVE_DI_11",   // "SENSOR"
              "SIMULACE_ON/OFF" := "SIMULACE",
              SIGNAL_OUT => #SEN_STRUCT.dvere_L_A,
              ENO => #_w3);
   #dvere_L_B(EN := #_w3,   // "SENSOR"
              SIGNAL_IN := "RESERVE_DI_12",
              "SIMULACE_ON/OFF" := "SIMULACE",
              SIGNAL_OUT => #SEN_STRUCT.dvere_L_B,
              ENO => #_w4);
   #dvere_P_A(EN := #_w4,   // "SENSOR"
              SIGNAL_IN := "RESERVE_DI_13",
              "SIMULACE_ON/OFF" := "SIMULACE",
              SIGNAL_OUT => #SEN_STRUCT.dvere_P_A,
              ENO => #_w5);
   IF #_w5 THEN
       #dvere_P_B(SIGNAL_IN := "RESERVE_DI_14",   // "SENSOR"
                  "SIMULACE_ON/OFF" := "SIMULACE",
                  SIGNAL_OUT => #SEN_STRUCT.dvere_P_B,
                  SIGNAL_OUT_NEG => #SEN_STRUCT.L1_NOT_OK);
   END_IF;
END_REGION

REGION Network 3 (SCL): ALARMY OP1/OP2 -> HMI
   // ===== ALARMY -> HMI (DB_ALARM.alarm_line, HMI ID 1-16) =====
   // bit 9 (ID 10 aplikator) a bit 14 (ID 15 tlak vzduchu) = firemni standard, nepouzivat

   // bit 0 - tiskarna nekomunikuje (OP2 se nevrati do kroku 5 do 15 s)
   "DB_ALARM".T_tiskarna.TON(IN := "AUTOMAT" AND "OP2_DB".SQCR <> 5,
                             PT := T#15S);
   "DB_ALARM".alarm_line.%X0 := "DB_ALARM".T_tiskarna.Q;

   // bity 1-3 - kamery offline (jen v automatu)
   "DB_ALARM".alarm_line.%X1 := "AUTOMAT" AND NOT "COG_FOLIE_L_is3800-Online";
   "DB_ALARM".alarm_line.%X2 := "AUTOMAT" AND NOT "COG_FOLIE_P_is3800-Online";
   "DB_ALARM".alarm_line.%X3 := "AUTOMAT" AND NOT "COG_ETIKETA_is3800-Online"
   AND NOT "OP1_DB".Kam_Etiketa_Job.aktivni;   // pri loadu jobu je kamera chvili offline

   // bit 4 - chybne datum v recepture
   "DB_ALARM".alarm_line.%X4 := "OP2_DB".Tisk.datum_chyba;

   // bit 5 - fronta plna
   "DB_ALARM".alarm_line.%X5 := "OP1_DB".Kamera.fronta_plna;

   // bit 6 - job horni kamery se nenacetl
   //"DB_ALARM".alarm_line.%X6 := "OP1_DB".Kam_Etiketa_Job.chyba;

   // bity 7-8 - otevrene dvere (signaly ze site "alarmy")
   "DB_ALARM".alarm_line.%X7 := "DB_ALARM".WRONG.dvere_L_tevreny;
   "DB_ALARM".alarm_line.%X8 := "DB_ALARM".WRONG.dvere_P_otevreny;

   // souhrnny alarm -> KA19 blika, HMI_ALARM = 10
   "alrm_global" := "DB_ALARM".alarm_line <> 0;
   "DB_ALARM".ALARM.ALARM_GLOBAL := "alrm_global";
END_REGION

